(* IEC 61131-3 sources: JingjiangArm/moonboxpro_arm_8.4/Application/Application/任务列表/ExtTask/动作处理/动作处理 (part 2) *)

(* ---- KS_FB_GrpFetchIOCtrl.st ---- *)
(*@CES
Name=KS_FB_GrpFetchIOCtrl
Type=FunctionBlock
TypeGuid=6f9dac99-8de1-4efc-8465-68ac443b7d08
Guid=a7ec576d-c0a8-4898-9e79-82769fd09b46
HasDeclaration=True
HasImplementation=True
*)
{DECLARATION}
FUNCTION_BLOCK KS_FB_GrpFetchIOCtrl
VAR_INPUT
	i_xEn: BOOL;
	i_iGrpId: INT;
	i_pstStEvtReq: POINTER TO StEvtReq; (* 沿触发标志 *)
	i_pstStSysCfgStruct: POINTER TO StSysCfgStruct;
	i_pastStIOMap_Main_FE						: POINTER TO ARRAY [1..4] OF StIOMap_Main_FE;(*轴io数据区域|AB系*)
	i_pastStIOMap_Axis_FE					: POINTER TO ARRAY [1..MAX_UNIT_NUM] OF StIOMap_Axis_FE;(*轴io数据区域|`````````````````````````````````````````````*)
	i_pastStIOMap_Axis_Extra_FE				: POINTER TO ARRAY [1..MAX_UNIT_NUM] OF StIOMap_Axis_Extra_FE;
	i_pastStIOMap_UwRw_FE_Uw					: POINTER TO ARRAY [1..2] OF StIOMap_UwRw_FE;(*轴io数据区域|AB系*)
	i_pastStIOMap_UwRw_FE_Rw					: POINTER TO ARRAY [1..2] OF StIOMap_UwRw_FE;(*轴io数据区域|AB系*)

	i_iUMax: INT;(*最大色组*)
	i_dwEquipmentProf: DWORD;(*机型：bit20:双收双放bit21:A放B收*)
	i_xUseRealStationOnRingnet: BOOL;(*使用真实站点*)
	i_axLinkage: ARRAY [1..MAX_UNIT_NUM] OF BOOL;
	i_axThisUnitEna: ARRAY [1..MAX_UNIT_NUM] OF BOOL;
	i_axSwitchOn_CoatingPrn: ARRAY [1..MAX_UNIT_NUM] OF BOOL;

	i_xIsValid_If_I: BOOL;
	i_xIsValid_If_II: BOOL;
	i_xIsValid_Of_I: BOOL;
	i_xIsValid_Of_II: BOOL;
//	i_pstStRingInfVer1: POINTER TO StRingInfVer1; (* 所有站点列表 *)

	//2026.5.20.133000 by liu.yt 使用map生成的系统站信息列表@根据实际站生成
	//i_pstStStationInfo_KS: POINTER TO StStationInfo_KS;
	(*输出列表*)
	i_pstStSysStationInf	: POINTER TO StSysStationInf;
	i_pxInit_StationList	: POINTER TO BOOL;

END_VAR
VAR_OUTPUT
	o_xEn: BOOL;
	o_iErNo: INT;
	o_iGrpAxisNum_Pu: INT; (* 系的色组数量|色组按照从小到大排序了 *)
	o_iGrpAxisTotalNum: INT; (* 系的轴数量 *)
	o_aiGrpAxisList: ARRAY [1..MAX_UNIT_NUM] OF INT; (* 系的轴列表 *)
	o_iIOGrpIdx_Uw: INT; (* 放料id *)
	o_iIOGrpIdx_Rw: INT; (* 收料id *)
	o_iAxisId_If_IOMapUse: INT; (* 放牵轴id *)
	o_iAxisId_Of_IOMapUse: INT; (* 收牵轴id *)
	o_aiGrpServoAxisList_Uw: ARRAY [1..2] OF INT := [2(-1)]; (* 2021.5.7.150202/目前仅支持双工位/[1]放置A轴/[2]放置B轴/轴id(-1)表无效 *)
	o_aiGrpServoAxisList_Rw: ARRAY [1..2] OF INT := [2(-1)]; (* 2021.5.7.150202/目前仅支持双工位/[1]放置A轴/[2]放置B轴/轴id(-1)表无效 *)

	(*2022.5.25.103645 增加联动轴*)
	o_iGrpLinkageAxisNum_Pu: INT; (* 系的色组联动轴数量|色组按照从小到大排序了 *)
	o_aiGrpLinkageAxisList: ARRAY [1..MAX_UNIT_NUM] OF INT; (* 系的联动轴列表 *)
	(*2023.09.04.131040 增加了色序列表的输出*)
	o_iGrpArcAxisNum_Pu: INT; (* 系的色联动轴套色打开数量|色组按照从小到大排序了 *)
	o_aiGrpArcAxisList: ARRAY [1..MAX_UNIT_NUM] OF INT; (* 系的联动轴套色打开列表 *)
	o_aiGrpArcIdList: ARRAY [1..MAX_UNIT_NUM] OF INT; (* 系的联动轴套色Id列表@2024.02.22.083346 套色id有可能会手动修改 *)
	o_aiGrpFollowArcIdList: ARRAY [1..MAX_UNIT_NUM] OF INT; (* 系的联动轴套色跟踪色序Id列表@2024.02.22.083346 和套色个数同步更新*)

(*运动列表*)
	o_iAxisNum_Trap: INT;(*点位运动轴数量*)
	o_aiStationList_Trap: ARRAY [1..MAX_STATION_NUM] OF INT;(*点位运动轴列表*)
	o_iAxisNum_Gear: INT;(*电子齿轮运动轴数量*)
	o_aiStationList_Gear: ARRAY [1..MAX_STATION_NUM] OF INT;(*电子齿轮运动轴列表*)
	o_iAxisNum_GantrayTrap: INT;(*龙门点位运动组数量*)
	o_aiStationList_GantrayTrap: ARRAY [1..MAX_STATION_NUM] OF INT;(*龙门点位运动轴列表*)
	o_iAxisNum_Jog: INT;(*龙门点位运动组数量*)
	o_aiStationList_Jog: ARRAY [1..MAX_STATION_NUM] OF INT;(*龙门点位运动轴列表*)
	o_iAxisNum_All: INT;
	o_aiStationList_All: ARRAY [1..MAX_STATION_NUM] OF INT;
	o_aiIndexList_All_Trap: ARRAY [1..MAX_STATION_NUM] OF INT;(*点位运动轴列表*)
	o_aiIndexList_All_Gear: ARRAY [1..MAX_STATION_NUM] OF INT;(*电子齿轮运动轴列表*)
	o_aiIndexList_All_Gantray: ARRAY [1..MAX_STATION_NUM] OF INT;(*龙门点位运动轴列表*)
	o_aiIndexList_All_Jog: ARRAY [1..MAX_STATION_NUM] OF INT;(*龙门点位运动轴列表*)
	o_axFlag_SlaveUseCmm_Pro: ARRAY [1..MAX_UNIT_NUM] OF BOOL;(*色组使用PRO/月光宝盒*)
	//2026.04.10.145314
	o_dwAxisFlags_Estop:DWORD;(*系急停状态*)
END_VAR
VAR_IN_OUT
	io_abyColorIdCurrent: ARRAY [1..MAX_UNIT_NUM] OF BYTE;(*色组色序*)
	io_abyFollowColorId: ARRAY [1..MAX_UNIT_NUM] OF BYTE;
END_VAR
VAR
	iN: INT;
	iK: INT;
	iTmpAxisId: INT;
	afbR_TRIG_EvtReq: ARRAY [1..17] OF R_TRIG; (* 上升沿触发器 *)
	dwMaskMonitoring_Estop: DWORD; (* 急停标志位输出 *)
	dwMaskMonitoring_Stop: DWORD;
	dwMaskMonitoring_FastStop: DWORD;
	dwMaskMonitoring_Tension: DWORD;
	dwMaskMonitoring_ManuSpdUp: DWORD;
	dwMaskMonitoring_ManuSpdDn: DWORD;
	dwMaskMonitoring_Ink: DWORD;
	dwMaskMonitoring_Prestart: DWORD;
	dwMaskMonitoring_PressAll: DWORD;
	dwMaskMonitoring_UnpressAll: DWORD;
	dwMaskMonitoring_Print: DWORD;
	dwMaskMonitoring_AlarmBell: DWORD;
	dwMaskMonitoring_AllInchRun: DWORD;
	dwMaskMonitoring_AllExhBlower: DWORD;
	dwMaskMonitoring_AllCoolBlower: DWORD;
	dwMaskMonitoring_AllHotBlower: DWORD;
	dwMaskMonitoring_AllHeating: DWORD;
	xIsDualUwRw: BOOL := FALSE; (* 双收双放 *)
	xAsOneMachine: BOOL := FALSE; (* A放B收结构 *)
	iUnitId: INT;
	iGrpId: INT;
	iTypeId: INT;
	iAxisTypeId: INT;
	xInit_ColorId: BOOL;(*开机初始化一次色序ID*)
	byColorID: BYTE;
	pstStIOMap_AxisBasic: POINTER TO StIOMap_Axis_FE; (* 基础io *)
	pstStIOMap_AxisExtra: POINTER TO StIOMap_Axis_Extra_FE; (* 扩展io *)
	axArcEnSts_Bak:ARRAY [1..MAX_STATION_NUM] OF BOOL;
	abyArcId_Bak:ARRAY [1..MAX_STATION_NUM] OF BYTE;
	iUnitId_Rd: INT;
	iTypeId_Rd: INT;
	//iAxisId_Rd: INT;
	//iCoreId_Rd: INT;
	//iGroupId_Rd: INT;
	//iAdjAxisId_Rd: INT;

	//2026.5.20.133421 by liu.yt
	pstStationInf:POINTER TO StStationInf;//每个站的信息
END_VAR

{IMPLEMENTATION}
o_xEn:= i_xEn;
o_iErNo:= 0;

(* 返回值初始化 *)
o_iIOGrpIdx_Uw:= -1; (* 放料io系id初始化 *)
o_iIOGrpIdx_Rw:= -1; (* 收料io系id初始化 *)
o_iAxisId_If_IOMapUse:= -1; (* 放牵轴id初始化 *)
o_iAxisId_Of_IOMapUse:= -1; (* 收牵轴id初始化 *)
o_iGrpAxisNum_Pu:= 0; (* 输出色组数量初始化 *)
o_iGrpAxisTotalNum:= 0; (* 输出总轴数量初始化 *)
o_iGrpLinkageAxisNum_Pu:= 0; (* 输出联动色组数量初始化 *)
o_iGrpArcAxisNum_Pu:=0;
FOR iN:=1 TO MAX_UNIT_NUM BY 1 DO(* 轴列表初始化 *)
	o_aiGrpAxisList[iN]:= -1;
	o_aiGrpLinkageAxisList[iN]:= -1;
	o_aiGrpArcAxisList[iN]:=-1;
	o_aiGrpArcIdList[iN]:=-1;(*2024.02.22.083413*)
	o_aiGrpFollowArcIdList[iN]:=-1;
END_FOR
o_aiGrpServoAxisList_Uw[1]:= -1;
o_aiGrpServoAxisList_Uw[2]:= -1;

o_aiGrpServoAxisList_Rw[1]:= -1;
o_aiGrpServoAxisList_Rw[2]:= -1;

(* 2018.9.4.162654\增加的监控初始化 *)
dwMaskMonitoring_Estop:= 0;
dwMaskMonitoring_Stop:= 0;
dwMaskMonitoring_Tension:= 0;
dwMaskMonitoring_ManuSpdUp:= 0;
dwMaskMonitoring_ManuSpdDn:= 0;
dwMaskMonitoring_Ink:= 0;
dwMaskMonitoring_Prestart:= 0;
dwMaskMonitoring_PressAll:= 0;
dwMaskMonitoring_UnpressAll:= 0;
dwMaskMonitoring_Print:= 0;
dwMaskMonitoring_AlarmBell:= 0;
dwMaskMonitoring_AllInchRun:= 0;
dwMaskMonitoring_AllExhBlower:= 0;
dwMaskMonitoring_AllCoolBlower:= 0;
dwMaskMonitoring_AllHotBlower:= 0;
dwMaskMonitoring_AllHeating:= 0;

IF i_xEn THEN
	IF (i_iGrpId=1 OR i_iGrpId=2) AND
		i_pstStEvtReq<>0 AND
		i_pastStIOMap_Main_FE<>0 AND
		i_pastStIOMap_Axis_FE<>0 AND
		i_pastStIOMap_Axis_Extra_FE<>0 AND
		i_pastStIOMap_UwRw_FE_Uw<>0 AND
		i_pastStIOMap_UwRw_FE_Rw<>0 AND
		i_pxInit_StationList<>0 THEN
		KS_InitStEvtReq(i_pstStEvtReq); (* 初始化StEvtReq@2018.7.31.094400 *)
		xIsDualUwRw:= i_dwEquipmentProf.20;
		xAsOneMachine:= i_dwEquipmentProf.21;
		IF NOT(i_iUMax>=1 AND i_iUMax<=16) THEN
			o_iErNo:=-4;
			RETURN;
		END_IF
		IF xIsDualUwRw AND xAsOneMachine AND i_iGrpId<>1 THEN(* A放B收\操作了A系以外的系 *)
			o_iErNo:= -2;
			RETURN;
		ELSIF (NOT xIsDualUwRw) AND i_iGrpId<>1 THEN(* 对于标准机型操作了A系以外的系 *)
			o_iErNo:= -3;
			RETURN;
		ELSE(* 其余正常情况 *)
			(* 生成当前系数的色组轴号列表|
			/*目前1个系内的放牵和收牵只认为各有1个,所以读取轴类型是牵引的会覆盖前面的取值 *)
			IF i_xUseRealStationOnRingnet THEN
// 				FOR iN:=1 TO i_pstStStationInfo_KS^.iStationNum BY 1 DO
// 					KS_GetAxisIdForMotByStation_V2(
// 						i_iStationId:= i_pstStStationInfo_KS^.aiStationId_List[iN],
// 						i_piAxisId:= ADR(iAxisId_Rd),
// 						i_piTypeId:= ADR(iTypeId_Rd),
// 						i_piUnitId:= ADR(iUnitId_Rd),
// 						i_piCoreId:= ADR(iCoreId_Rd),
// 						i_piGroupId:= ADR(iGroupId_Rd),
// 						i_piAdjAxisId:= ADR(iAdjAxisId_Rd),
// 						i_pstStSysStationInf:= ADR(g_stStSysStationInf));
// 					IF iUnitId_Rd>=1 AND iUnitId<=MAX_UNIT_NUM THEN
// 						iGrpId:= KS_GetGrpIdByAxisId(iUnitId,ADR(g_stStSysParam),ADR(iAxisTypeId));
// 						//2026.5.12.112929就用版辊驱动器数量输出轴列表吧
// 						IF iGrpId= i_iGrpId THEN
// 							IF iTypeId_Rd=TYPE_UNIT_PRN THEN
// 								o_iGrpAxisNum_Pu:= o_iGrpAxisNum_Pu+1;
// 								o_aiGrpAxisList[o_iGrpAxisNum_Pu]:= iUnitId_Rd;
// 							END_IF
// 						END_IF
// 					END_IF
// 				END_FOR
				//2026.5.20.133216 by liu.yt 重新生成列表@根据实际站
				FOR iN:=1 TO BYTE_TO_INT(i_pstStSysStationInf^.byStationNum) BY 1 DO
					pstStationInf:=ADR(i_pstStSysStationInf^.astStationInf[iN]);

					KS_GetAxisIdForMotByStation_V2(
						i_iStationId:= pstStationInf^.iStationId,
						i_piAxisId:= 0,
						i_piTypeId:= ADR(iTypeId_Rd),
						i_piUnitId:= ADR(iUnitId_Rd),
						i_piCoreId:= 0,
						i_piGroupId:= 0,
						i_piAdjAxisId:= 0,
						i_pstStSysStationInf:= i_pstStSysStationInf);
					IF iUnitId_Rd>=1 AND iUnitId_Rd<=MAX_UNIT_NUM THEN//色组id合法@1个色组可能会存在多个不同功能站号返回。我们只检查色组轴
						iGrpId:= KS_GetGrpIdByAxisId(iUnitId_Rd,ADR(g_stStSysParam),ADR(iAxisTypeId));
						//2026.5.12.112929就用版辊驱动器数量输出轴列表吧
						IF iGrpId= i_iGrpId THEN
							IF iTypeId_Rd=TYPE_UNIT_CTL THEN
								o_iGrpAxisNum_Pu:= o_iGrpAxisNum_Pu+1;
								o_aiGrpAxisList[o_iGrpAxisNum_Pu]:= iUnitId_Rd;
							END_IF
						END_IF
					END_IF
				END_FOR
			ELSE
				(* 2020.9.11.134731
				** 按照系统配置的色组填充列表|
				** *)
				FOR iUnitId:=1 TO i_iUMax BY 1 DO
					o_iGrpAxisNum_Pu:= o_iGrpAxisNum_Pu+1;
					o_aiGrpAxisList[o_iGrpAxisNum_Pu]:= iUnitId;
				END_FOR
			END_IF

			(* **
			** 将牵引轴使能出来@2019.4.26.171841
			** 针对给了使能|但没有给牵引指定一个有效的轴id
			** *)
			IF NOT xIsDualUwRw THEN(* 非双收双放 *)
				(* 放牵轴id *)
				IF i_xIsValid_If_I THEN
					o_iAxisId_If_IOMapUse:= 1;
				END_IF

				(* 收牵轴id *)
				IF i_xIsValid_Of_I THEN
					o_iAxisId_Of_IOMapUse:= 2;
				END_IF
			ELSE(* 双收双放 *)
				IF xAsOneMachine THEN(* A放B收 *)
					IF i_iGrpId=1 THEN
						(* 放牵轴id *)
						IF i_xIsValid_If_I THEN
							o_iAxisId_If_IOMapUse:= 1;
						END_IF

						(* 收牵轴id *)
						IF i_xIsValid_Of_II THEN
							o_iAxisId_Of_IOMapUse:= 4;
						END_IF
					END_IF
				ELSE(* A放A收|B放B收 *)
					IF i_iGrpId=1 THEN
						(* 放牵轴id *)
						IF i_xIsValid_If_I THEN
							o_iAxisId_If_IOMapUse:= 1;
						END_IF

						(* 收牵轴id *)
						IF i_xIsValid_Of_I THEN
							o_iAxisId_Of_IOMapUse:= 2;
						END_IF
					ELSE(* B系 *)
						(* 放牵轴id *)
						IF i_xIsValid_If_II THEN
							o_iAxisId_If_IOMapUse:= 3;
						END_IF

						(* 收牵轴id *)
						IF i_xIsValid_Of_II THEN
							o_iAxisId_Of_IOMapUse:= 4;
						END_IF
					END_IF
				END_IF
			END_IF
			(* 色组按从小到大的编号排列 *)
			FOR iN:=o_iGrpAxisNum_Pu TO 2 BY -1 DO
				FOR iK:=1 TO iN BY 1 DO
					IF o_aiGrpAxisList[iN]<o_aiGrpAxisList[iK] THEN
						iTmpAxisId:= o_aiGrpAxisList[iN];
						o_aiGrpAxisList[iN]:= o_aiGrpAxisList[iK];
						o_aiGrpAxisList[iK]:= iTmpAxisId;
					END_IF
				END_FOR
			END_FOR

			(* 在色组轴号之后追加牵引轴编号 *)
			o_iGrpAxisTotalNum:= o_iGrpAxisNum_Pu;
(*2026.5.12.132915这个列表只放色组相关的
			(* 放牵 *)
			IF o_iAxisId_If_IOMapUse>=1 AND o_iAxisId_If_IOMapUse<=MAX_STATION_NUM THEN
				o_iGrpAxisTotalNum:= o_iGrpAxisTotalNum+1;
				o_aiGrpAxisList[o_iGrpAxisTotalNum]:= o_iAxisId_If_IOMapUse;
			END_IF

			(* 收牵 *)
			IF o_iAxisId_Of_IOMapUse>=1 AND o_iAxisId_Of_IOMapUse<=MAX_STATION_NUM THEN
				o_iGrpAxisTotalNum:= o_iGrpAxisTotalNum+1;
				o_aiGrpAxisList[o_iGrpAxisTotalNum]:= o_iAxisId_Of_IOMapUse;
			END_IF
*)
			(*2022.5.25.104049 增加联动轴的列表输出*)
			FOR iN:=1 TO o_iGrpAxisNum_Pu BY 1 DO
				iTmpAxisId:= o_aiGrpAxisList[iN];
				IF iTmpAxisId>0 THEN
					IF i_axLinkage[iTmpAxisId] THEN(*联动*)
						o_iGrpLinkageAxisNum_Pu:=o_iGrpLinkageAxisNum_Pu+1;
						o_aiGrpLinkageAxisList[o_iGrpLinkageAxisNum_Pu]:=iTmpAxisId;
					END_IF
				END_IF
			END_FOR

			(*2023.09.04.131214 增加联动轴套色打开的列表输出*)
			IF xInit_ColorId THEN
				FOR iN:=1 TO o_iGrpLinkageAxisNum_Pu BY 1 DO
					iTmpAxisId:= o_aiGrpLinkageAxisList[iN];
					IF iTmpAxisId>0 THEN
						IF io_abyColorIdCurrent[iTmpAxisId]>0 AND io_abyColorIdCurrent[iTmpAxisId]<=MAX_UNIT_NUM THEN(*色序合法*)
							o_iGrpArcAxisNum_Pu:=o_iGrpArcAxisNum_Pu+1;
							o_aiGrpArcAxisList[o_iGrpArcAxisNum_Pu]:=iTmpAxisId;
							o_aiGrpArcIdList[o_iGrpArcAxisNum_Pu]:=io_abyColorIdCurrent[iTmpAxisId];(*2024.02.22.083448 套色id也统计出来*)
							o_aiGrpFollowArcIdList[o_iGrpArcAxisNum_Pu]:=io_abyFollowColorId[iTmpAxisId];(*2024.02.22.112812 界面修改或者一些开关控制*)
						END_IF
					END_IF
				END_FOR
			END_IF

			IF xIsDualUwRw THEN
				(* 双收双放 *)

				IF xAsOneMachine THEN
					(* A放B收 *)
					o_iIOGrpIdx_Uw:= 1;
					o_iIOGrpIdx_Rw:= 2;
				ELSE
					(* A/B系各自用各自的 *)
					IF i_iGrpId=1 THEN
						o_iIOGrpIdx_Uw:= 1;
						o_iIOGrpIdx_Rw:= 1;
					ELSE
						o_iIOGrpIdx_Uw:= 2;
						o_iIOGrpIdx_Rw:= 2;
					END_IF
				END_IF
			ELSE(* 普通机型\只看A系 *)
				o_iIOGrpIdx_Uw:= 1;
				o_iIOGrpIdx_Rw:= 1;
			END_IF

			(* 放料和收料的急停按钮 *)
			IF i_pastStIOMap_UwRw_FE_Uw^[o_iIOGrpIdx_Uw].i_xEstop THEN(* 放料急停 *)
				dwMaskMonitoring_Estop:= dwMaskMonitoring_Estop OR SHL(DWORD#1,20);
				i_pstStEvtReq^.xEvt_Estop:= TRUE;
			END_IF
			IF i_pastStIOMap_UwRw_FE_Rw^[o_iIOGrpIdx_Rw].i_xEstop THEN(* 收料急停 *)
				dwMaskMonitoring_Estop:= dwMaskMonitoring_Estop OR SHL(DWORD#1,21);
				i_pstStEvtReq^.xEvt_Estop:= TRUE;
			END_IF

			(*放牵收牵的按钮处理*)
			IF i_pastStIOMap_Main_FE^[o_iAxisId_If_IOMapUse].i_xEstop OR
				i_pastStIOMap_Main_FE^[o_iAxisId_Of_IOMapUse].i_xEstop THEN
				i_pstStEvtReq^.xEvt_Estop:= TRUE;
			END_IF
			IF i_pastStIOMap_Main_FE^[o_iAxisId_If_IOMapUse].i_xStop OR
				i_pastStIOMap_Main_FE^[o_iAxisId_Of_IOMapUse].i_xStop THEN
				i_pstStEvtReq^.xEvt_Stop:= TRUE;
			END_IF
			IF i_pastStIOMap_Main_FE^[o_iAxisId_If_IOMapUse].i_xFastStop OR
				i_pastStIOMap_Main_FE^[o_iAxisId_Of_IOMapUse].i_xFastStop THEN
				//2026.06.04.145510 变量写错了 by liu.yt
				//i_pstStEvtReq^.xEvt_Stop:= TRUE;
				i_pstStEvtReq^.xEvt_FastStop:= TRUE;
			END_IF
			IF i_pastStIOMap_Main_FE^[o_iAxisId_If_IOMapUse].i_xTension OR
				i_pastStIOMap_Main_FE^[o_iAxisId_Of_IOMapUse].i_xTension THEN
				i_pstStEvtReq^.xEvt_Tension:= TRUE;
			END_IF
			IF i_pastStIOMap_Main_FE^[o_iAxisId_If_IOMapUse].i_xAcc OR
				i_pastStIOMap_Main_FE^[o_iAxisId_Of_IOMapUse].i_xAcc THEN
				i_pstStEvtReq^.xEvt_ManuSpdUp:= TRUE;
			END_IF
			IF i_pastStIOMap_Main_FE^[o_iAxisId_If_IOMapUse].i_xDec OR
				i_pastStIOMap_Main_FE^[o_iAxisId_Of_IOMapUse].i_xDec THEN
				i_pstStEvtReq^.xEvt_ManuSpdDn:= TRUE;
			END_IF
			IF i_pastStIOMap_Main_FE^[o_iAxisId_If_IOMapUse].i_xInk OR
				i_pastStIOMap_Main_FE^[o_iAxisId_Of_IOMapUse].i_xInk THEN
				i_pstStEvtReq^.xEvt_Ink:= TRUE;
			END_IF
			IF i_pastStIOMap_Main_FE^[o_iAxisId_If_IOMapUse].i_xPrestart OR
				i_pastStIOMap_Main_FE^[o_iAxisId_Of_IOMapUse].i_xPrestart THEN
				i_pstStEvtReq^.xEvt_Prestart:= TRUE;
			END_IF
			IF i_pastStIOMap_Main_FE^[o_iAxisId_If_IOMapUse].i_xPrint OR
				i_pastStIOMap_Main_FE^[o_iAxisId_Of_IOMapUse].i_xPrint THEN
				i_pstStEvtReq^.xEvt_Print:= TRUE;
			END_IF
			IF i_pastStIOMap_Main_FE^[o_iAxisId_If_IOMapUse].i_xPressAll OR
				i_pastStIOMap_Main_FE^[o_iAxisId_Of_IOMapUse].i_xPressAll THEN
				i_pstStEvtReq^.xEvt_PressAll:= TRUE;
			END_IF
			IF i_pastStIOMap_Main_FE^[o_iAxisId_If_IOMapUse].i_xUnPressAll OR
				i_pastStIOMap_Main_FE^[o_iAxisId_Of_IOMapUse].i_xUnPressAll THEN
				i_pstStEvtReq^.xEvt_UnPressAll:= TRUE;
			END_IF
			IF i_pastStIOMap_Main_FE^[o_iAxisId_If_IOMapUse].i_xAlarmBell OR
				i_pastStIOMap_Main_FE^[o_iAxisId_Of_IOMapUse].i_xAlarmBell THEN
				i_pstStEvtReq^.xEvt_AlarmBell:= TRUE;
			END_IF

			IF i_pastStIOMap_Main_FE^[o_iAxisId_If_IOMapUse].i_xAllExhBlower_Up OR
				i_pastStIOMap_Main_FE^[o_iAxisId_Of_IOMapUse].i_xAllExhBlower_Up OR
				i_pastStIOMap_Main_FE^[o_iAxisId_If_IOMapUse].i_xAllExhBlower_Dn OR
				i_pastStIOMap_Main_FE^[o_iAxisId_Of_IOMapUse].i_xAllExhBlower_Dn THEN
				(* 整机排风 *)
				i_pstStEvtReq^.xEvt_AllExhBlower:= TRUE;
			END_IF

			IF i_pastStIOMap_Main_FE^[o_iAxisId_If_IOMapUse].i_xAllCoolBlower OR
				i_pastStIOMap_Main_FE^[o_iAxisId_Of_IOMapUse].i_xAllCoolBlower THEN
				(* 整机冷风 *)
				i_pstStEvtReq^.xEvt_AllCoolBlower:= TRUE;
			END_IF
			IF i_pastStIOMap_Main_FE^[o_iAxisId_If_IOMapUse].i_xAllHotBlower OR
				i_pastStIOMap_Main_FE^[o_iAxisId_Of_IOMapUse].i_xAllHotBlower THEN
				(* 整机热风 *)
				i_pstStEvtReq^.xEvt_AllHotBlower:= TRUE;
			END_IF
			IF i_pastStIOMap_Main_FE^[o_iAxisId_If_IOMapUse].i_xAllHeating OR
				i_pastStIOMap_Main_FE^[o_iAxisId_Of_IOMapUse].i_xAllHeating THEN
				(* 整机加热 *)
				i_pstStEvtReq^.xEvt_AllHeating:= TRUE;
			END_IF

			(* 默认3档开关 作互斥 *)
			IF i_pastStIOMap_Main_FE^[o_iAxisId_Of_IOMapUse].i_xTapPosition_Breaking THEN(* 2018.7.16.151749\断料档位 *)
				i_pstStEvtReq^.xEvt_TapPosition_Breaking:= TRUE;
				i_pstStEvtReq^.xEvt_TapPosition_UniformInk:= FALSE;
				i_pstStEvtReq^.xEvt_TapPosition_Printing:= FALSE;
			ELSIF i_pastStIOMap_Main_FE^[o_iAxisId_Of_IOMapUse].i_xTapPosition_UniformInk THEN(* 2018.7.16.152023\匀墨档位 *)
				i_pstStEvtReq^.xEvt_TapPosition_UniformInk:= TRUE;
				i_pstStEvtReq^.xEvt_TapPosition_Breaking:= FALSE;
				i_pstStEvtReq^.xEvt_TapPosition_Printing:= FALSE;
			ELSE(* 2018.7.16.152128\印刷档位 *)
				i_pstStEvtReq^.xEvt_TapPosition_Printing:= TRUE;
				i_pstStEvtReq^.xEvt_TapPosition_Breaking:= FALSE;
				i_pstStEvtReq^.xEvt_TapPosition_UniformInk:= FALSE;
			END_IF

			(* 影响整机的逻辑按钮\所有轴上可能都有\就在FOR循环里面检查(当然要包含牵引) *)
			byColorID:=0;(*2022.6.8.101746*)
			FOR iN:=1 TO o_iGrpAxisNum_Pu BY 1 DO
				iUnitId:= o_aiGrpAxisList[iN]; (* 列表由于本地生成\所以iAxisId可以不检查 *)
				pstStIOMap_AxisBasic:= ADR(i_pastStIOMap_Axis_FE^[iUnitId]); (* 基础io表 *)
				pstStIOMap_AxisExtra:= ADR(i_pastStIOMap_Axis_Extra_FE^[iUnitId]); (* 扩展io表 *)

				IF pstStIOMap_AxisBasic^.i_xEstop THEN
					(* 急停 *)
					i_pstStEvtReq^.xEvt_Estop:= TRUE;
					dwMaskMonitoring_Estop:= dwMaskMonitoring_Estop OR SHL(DWORD#1,iUnitId-1);
				END_IF
				IF pstStIOMap_AxisBasic^.i_xStop THEN
					(* 停机 *)
					i_pstStEvtReq^.xEvt_Stop:= TRUE;
					dwMaskMonitoring_Stop:= dwMaskMonitoring_Stop OR SHL(DWORD#1,iUnitId-1);
				END_IF

				IF pstStIOMap_AxisBasic^.i_xAcc THEN
					(* 手动加速 *)
					i_pstStEvtReq^.xEvt_ManuSpdUp:= TRUE;
					dwMaskMonitoring_ManuSpdUp:= dwMaskMonitoring_ManuSpdUp OR SHL(DWORD#1,iUnitId-1);
				END_IF
				IF pstStIOMap_AxisBasic^.i_xDec THEN
					(* 手动减速 *)
					i_pstStEvtReq^.xEvt_ManuSpdDn:= TRUE;
					dwMaskMonitoring_ManuSpdDn:= dwMaskMonitoring_ManuSpdDn OR SHL(DWORD#1,iUnitId-1);
				END_IF

				IF pstStIOMap_AxisBasic^.i_xAlarmBell THEN
					(* 警铃 *)
					i_pstStEvtReq^.xEvt_AlarmBell:= TRUE;
					dwMaskMonitoring_AlarmBell:= dwMaskMonitoring_AlarmBell OR SHL(DWORD#1,iUnitId-1);
				END_IF
				IF pstStIOMap_AxisBasic^.i_xInch AND
					i_axLinkage[iUnitId] THEN
					(* 整机单运行 *)
					i_pstStEvtReq^.xEvt_AllInchRun:= TRUE;
					dwMaskMonitoring_AllInchRun:= dwMaskMonitoring_AllInchRun OR SHL(DWORD#1,iUnitId-1);
				END_IF
			END_FOR

			//2026.5.9.172930
			//2026.04.10.145142 + 系急停变量赋值
			o_dwAxisFlags_Estop:=dwMaskMonitoring_Estop;

			(*2024.02.21.084550 优化套色id逻辑*)
			KS_GetArcIdList(
				TRUE(*i_xEn*),
				o_iGrpAxisNum_Pu(*i_iGrpAxisNum_Pu*),
				o_aiGrpAxisList(*i_aiGrpAxisList*),
				ADR(axArcEnSts_Bak)(*i_paxArcEnSts_Bak*),
				ADR(abyArcId_Bak)(*i_pabyArcId_Bak*),
				0(*i_piGrpArcAxisNum_Pu*),
				i_axLinkage,
				i_axThisUnitEna,
				i_axSwitchOn_CoatingPrn,
				ADR(io_abyColorIdCurrent));
			xInit_ColorId:=TRUE;

		END_IF

		(*2025.6.16.165421运动所有的轴列表处理一下*)
		IF NOT i_pxInit_StationList^ THEN
			i_pxInit_StationList^:= TRUE;
			o_iAxisNum_Trap:= 0;
			o_iAxisNum_Gear:= 0;
			o_iAxisNum_GantrayTrap:= 0;
			o_iAxisNum_Jog:= 0;
			o_iAxisNum_All:= 0;
			FOR iN:=1 TO MAX_STATION_NUM BY 1 DO
				o_aiStationList_Trap[iN]:= 0;
				o_aiStationList_Gear[iN]:= 0;
				o_aiStationList_GantrayTrap[iN]:= 0;
				o_aiStationList_All[iN]:= 0;
				o_aiIndexList_All_Trap[iN]:= 0;
				o_aiIndexList_All_Gear[iN]:= 0;
				o_aiIndexList_All_Gantray[iN]:= 0;
			END_FOR

			FOR iN:=1 TO i_pstStSysStationInf^.byStationNum BY 1 DO
				pstStationInf:=ADR(i_pstStSysStationInf^.astStationInf[iN]);
				KS_GetUnitIdAndTypeByStationId(
					pstStationInf^.iStationId ,//i_pstStRingInfVer1^.m_station_id_list[iN],//i_pstStStationInfo_KS^.aiStationId_List[iN], //,
					ADR(iUnitId),
					ADR(iTypeId),
					i_pstStSysCfgStruct);
				IF iTypeId= OBJ_IS_HORIZ_MOTION OR
					 iTypeId=OBJ_IS_PHOTOCELL THEN(*光电眼行走机构 | 2024.04.01.092649*)
					o_iAxisNum_Trap:= o_iAxisNum_Trap+1;
					IF o_iAxisNum_Trap<>0 THEN
						o_aiStationList_Trap[o_iAxisNum_Trap]:= pstStationInf^.iStationId;//i_pstStRingInfVer1^.m_station_id_list[iN];//
						o_aiIndexList_All_Trap[o_iAxisNum_Trap]:= iN;
					END_IF
				ELSIF iTypeId= OBJ_IS_PRN_ROLLER_PRESSURE_M OR
					iTypeId= OBJ_IS_PRN_ROLLER_PRESSURE_G OR
					iTypeId= OBJ_IS_NET_ROLLER_PRESSURE_M OR
					iTypeId= OBJ_IS_NET_ROLLER_PRESSURE_G OR
					iTypeId= OBJ_IS_STR_ROLLER_PRESSURE_M OR
					iTypeId= OBJ_IS_STR_ROLLER_PRESSURE_G THEN
					o_iAxisNum_GantrayTrap:= o_iAxisNum_GantrayTrap+1;
					IF o_iAxisNum_GantrayTrap<>0 THEN
						o_aiStationList_GantrayTrap[o_iAxisNum_GantrayTrap]:= pstStationInf^.iStationId;//i_pstStRingInfVer1^.m_station_id_list[iN];//;
						o_aiIndexList_All_Gantray[o_iAxisNum_GantrayTrap]:= iN;

					END_IF
				ELSIF iTypeId= OBJ_IS_UNWIND_A OR
					iTypeId= OBJ_IS_UNWIND_B OR
					iTypeId= OBJ_IS_REWIND_A OR
					iTypeId= OBJ_IS_REWIND_B OR
					iTypeId= OBJ_IS_INFEED OR
					iTypeId= OBJ_IS_OUTFEED OR
					iTypeId= OBJ_IS_BOTTOM_ROLLER OR
					iTypeId= OBJ_IS_PRN_ROLLER OR
					iTypeId= OBJ_IS_NET_ROLLER OR
					iTypeId= OBJ_IS_CENTRAL_DRUM THEN
					o_iAxisNum_Gear:= o_iAxisNum_Gear+1;
					IF o_iAxisNum_Gear<>0 THEN
						o_aiStationList_Gear[o_iAxisNum_Gear]:= pstStationInf^.iStationId;//i_pstStRingInfVer1^.m_station_id_list[iN];//;
						o_aiIndexList_All_Gear[o_iAxisNum_Gear]:= iN;

					END_IF

					//2026.05.08.141028 | + | 增加收放料伺服的标志
					IF iTypeId= OBJ_IS_UNWIND_A OR
						iTypeId= OBJ_IS_UNWIND_B OR
						iTypeId= OBJ_IS_REWIND_A OR
						iTypeId= OBJ_IS_REWIND_B THEN
						g_xUwRwIsServo := TRUE;
					END_IF
				//这部分的代码处理会有问题@2026.5.20.140553 by liu.yt
				ELSIF pstStationInf^.iStationId>=1
					AND pstStationInf^.iStationId<16
					AND (pstStationInf^.udiStationType=HY_YTPE_CMM_CR_PRO
					OR	pstStationInf^.udiStationType=HY_YTPE_CMM_CR) THEN//色组使用月光宝盒/PRO通讯
					IF pstStationInf^.udiStationType=HY_YTPE_CMM_CR_PRO THEN
						o_axFlag_SlaveUseCmm_Pro[pstStationInf^.iStationId]:= TRUE;
					ELSE
						o_axFlag_SlaveUseCmm_Pro[pstStationInf^.iStationId]:= FALSE;
					END_IF
				END_IF
				IF iTypeId= OBJ_IS_HORIZ_MOTION OR
					iTypeId= OBJ_IS_PRN_ROLLER_PRESSURE_M OR
					iTypeId= OBJ_IS_PRN_ROLLER_PRESSURE_G OR
					iTypeId= OBJ_IS_NET_ROLLER_PRESSURE_M OR
					iTypeId= OBJ_IS_NET_ROLLER_PRESSURE_G OR
					iTypeId= OBJ_IS_UNWIND_A OR
					iTypeId= OBJ_IS_UNWIND_B OR
					iTypeId= OBJ_IS_REWIND_A OR
					iTypeId= OBJ_IS_REWIND_B OR
					iTypeId= OBJ_IS_INFEED OR
					iTypeId= OBJ_IS_OUTFEED OR
					iTypeId= OBJ_IS_BOTTOM_ROLLER OR
					iTypeId= OBJ_IS_PRN_ROLLER OR
					iTypeId= OBJ_IS_NET_ROLLER OR
					iTypeId= OBJ_IS_CENTRAL_DRUM OR//所有参与运动的轴个数
					iTypeId= OBJ_IS_PHOTOCELL OR
					iTypeId= OBJ_IS_STR_ROLLER_PRESSURE_M OR
					iTypeId= OBJ_IS_STR_ROLLER_PRESSURE_G THEN//所有参与运动的轴个数
					o_iAxisNum_All:= o_iAxisNum_All+1;
					IF o_iAxisNum_All<>0 THEN
						o_aiStationList_All[o_iAxisNum_All]:= pstStationInf^.iStationId;//i_pstStRingInfVer1^.m_station_id_list[iN];//;
					END_IF
				END_IF
			END_FOR
		END_IF

		(*-----------end--------------------------*)

		(* 上升沿检测 *)
		afbR_TRIG_EvtReq[1](CLK:= i_pstStEvtReq^.xEvt_Estop, Q=> i_pstStEvtReq^.xReqEstop); (* 急停 *)
		afbR_TRIG_EvtReq[2](CLK:= i_pstStEvtReq^.xEvt_Stop, Q=> i_pstStEvtReq^.xReqStop); (* 停机 *)
		afbR_TRIG_EvtReq[3](CLK:= i_pstStEvtReq^.xEvt_Tension, Q=> i_pstStEvtReq^.xReqTension); (* 张力投入 *)
		afbR_TRIG_EvtReq[4](CLK:= i_pstStEvtReq^.xEvt_ManuSpdUp, Q=> i_pstStEvtReq^.xReqManuSpdUp); (* 手动加速|按着才加速 *)
		afbR_TRIG_EvtReq[5](CLK:= i_pstStEvtReq^.xEvt_ManuSpdDn, Q=> i_pstStEvtReq^.xReqManuSpdDn); (* 手动减速|按着才减速 *)
		afbR_TRIG_EvtReq[6](CLK:= i_pstStEvtReq^.xEvt_Ink, Q=> i_pstStEvtReq^.xReqInk); (* 空转 *)
		afbR_TRIG_EvtReq[7](CLK:= i_pstStEvtReq^.xEvt_Prestart, Q=> i_pstStEvtReq^.xReqPrestart); (* 启动|预备 *)
		afbR_TRIG_EvtReq[8](CLK:= i_pstStEvtReq^.xEvt_PressAll, Q=> i_pstStEvtReq^.xReqPressAll); (* 全体合压 *)
		afbR_TRIG_EvtReq[9](CLK:= i_pstStEvtReq^.xEvt_UnpressAll, Q=> i_pstStEvtReq^.xReqUnpressAll); (* 全体离压 *)
		afbR_TRIG_EvtReq[10](CLK:= i_pstStEvtReq^.xEvt_Print, Q=> i_pstStEvtReq^.xReqPrint); (* 印刷|联动 *)
		afbR_TRIG_EvtReq[11](CLK:= i_pstStEvtReq^.xEvt_AlarmBell, Q=> i_pstStEvtReq^.xReqAlarmBell); (* 警铃|按着才响 *)
		afbR_TRIG_EvtReq[12](CLK:= i_pstStEvtReq^.xEvt_AllInchRun, Q=> i_pstStEvtReq^.xReqAllInchRun); (* 整机单运行 *)
		afbR_TRIG_EvtReq[13](CLK:= i_pstStEvtReq^.xEvt_AllExhBlower, Q=> i_pstStEvtReq^.xReqAllExhBlower); (* 排风启动 *)
		afbR_TRIG_EvtReq[14](CLK:= i_pstStEvtReq^.xEvt_AllCoolBlower, Q=> i_pstStEvtReq^.xReqAllCoolBlower); (* 冷风启动 *)
		afbR_TRIG_EvtReq[15](CLK:= i_pstStEvtReq^.xEvt_AllHotBlower, Q=> i_pstStEvtReq^.xReqAllHotBlower); (* 热风启动 *)
		afbR_TRIG_EvtReq[16](CLK:= i_pstStEvtReq^.xEvt_AllHeating, Q=> i_pstStEvtReq^.xReqAllHeating); (* 加热启动 *)
		afbR_TRIG_EvtReq[17](CLK:= i_pstStEvtReq^.xEvt_FastStop, Q=> i_pstStEvtReq^.xReqFastStop); (* 快停按钮 *)
		(*记录日志和变频报警处理稍后*)
	END_IF
END_IF

(* ---- KS_FB_GrpIndicatorLampCtrl.st ---- *)
(*@CES
Name=KS_FB_GrpIndicatorLampCtrl
Type=FunctionBlock
TypeGuid=6f9dac99-8de1-4efc-8465-68ac443b7d08
Guid=046cf0cb-05a3-4565-9599-869039b6c2cc
HasDeclaration=True
HasImplementation=True
*)
{DECLARATION}
FUNCTION_BLOCK KS_FB_GrpIndicatorLampCtrl
VAR_INPUT
	i_xEn: BOOL;
	i_iGrpId:INT;
	i_iCustomerNameId:INT;
	i_iGrpAxisNum_PU: INT;
	i_aiGrpAxisList: ARRAY [1..MAX_UNIT_NUM] OF INT;
	i_pstStSysParam: POINTER TO StSysParam;
	i_pastStIOMap_AxisBasic: POINTER TO ARRAY [1..MAX_UNIT_NUM] OF StIOMap_Axis_FE;
	i_pastStIOMap_Main: POINTER TO ARRAY [1..4] OF StIOMap_Main_FE;(*基础io|*)
	i_iAxisId_If: INT;
	i_iAxisId_Of: INT;
END_VAR
VAR_OUTPUT
	o_xEno: BOOL;
	o_iErNo: INT;
END_VAR
VAR
	iN: INT;
	iAxisId: INT;
	pstStIOMap_AxisBasic: POINTER TO StIOMap_Axis_FE;
	pstStIOMap_Main: POINTER TO StIOMap_Main_FE;
	pstStIOMap_Main_If: POINTER TO StIOMap_Main_FE;
	pstStIOMap_Main_Of: POINTER TO StIOMap_Main_FE;
	tmNow: TIME;
	tmLastStateChanged_print: TIME;
	tmLastStateChanged_prestart: TIME; (* 2021.3.3.113856/上次状态改变的时间 *)
	tmLastStateChanged_Stop: TIME; (* 2022.4.10.001512/上次状态改变的时间 *)
	xLamp_Stop: BOOL;(*停止灯指示*)
END_VAR

{IMPLEMENTATION}
o_xEno:= i_xEn;
o_iErNo:= 0;
IF i_xEn THEN
	IF (i_iGrpAxisNum_PU>=0 AND i_iGrpAxisNum_PU<=MAX_UNIT_NUM) AND(*色组有效|*)
		i_pastStIOMap_AxisBasic<>0 THEN(*轴IO有效|*)

		tmNow:= TIME(); (* 2021.3.3.114019/ *)

		(*2022.4.9.225300 增加了停止时候停止指示灯的闪烁指示*)
		IF i_pstStSysParam^.astStGrpParam_UnSave[i_iGrpId].xFlag_Stoping  (*OR (*停止中|*)
			 i_pstStGrpParam^.xFlag_FastStoping*) THEN(*快速停止中*)
			IF tmNow-tmLastStateChanged_Stop>=T#200MS THEN
				xLamp_Stop:=NOT xLamp_Stop;(**)
				tmLastStateChanged_Stop:= tmNow; (* 2021.3.3.114723/ *)
			END_IF
		ELSE
			xLamp_Stop:=i_pstStSysParam^.astStGrpParam_UnSave[i_iGrpId].xFlag_Stop;
			tmLastStateChanged_Stop:= tmNow; (* 2021.3.3.114723/ *)
		END_IF

		FOR iN:=1 TO i_iGrpAxisNum_PU BY 1 DO
			iAxisId:= i_aiGrpAxisList[iN];
			IF iAxisId>=1 AND iAxisId<=MAX_UNIT_NUM THEN
				pstStIOMap_AxisBasic:=ADR(i_pastStIOMap_AxisBasic^[iAxisId]);(*读取轴IO|*)
				//pstStIOMap_Main_If:=ADR(i_pastStIOMap_Main^[i_iAxisId_If]);(*读取牵引轴IO|*)
				//pstStIOMap_Main_Of:=ADR(i_pastStIOMap_Main^[i_iAxisId_Of]);(*读取牵引轴IO|*)
				pstStIOMap_AxisBasic^.o_xLamp_Estop:= i_pstStSysParam^.astStGrpParam_UnSave[i_iGrpId].xFlag_Estop AND pstStIOMap_AxisBasic^.i_xEstop;(*急停灯输出|*)
				pstStIOMap_AxisBasic^.o_xLamp_Stop:= xLamp_Stop OR
												(NOT i_pstStSysParam^.astStUnitParam_Save[iAxisId].xLinkage AND NOT i_pstStSysParam^.astStGrpParam_UnSave[i_iGrpId].xFlag_Estop);(*停止灯输出|*)
				pstStIOMap_AxisBasic^.o_xLamp_Inch:= (i_pstStSysParam^.astStGrpParam_UnSave[i_iGrpId].xFlag_Ink OR i_pstStSysParam^.astStGrpParam_UnSave[i_iGrpId].xFlag_Print) AND (i_pstStSysParam^.astStUnitParam_Save[iAxisId].xLinkage);(*联动状态下空转或印刷|*)
				pstStIOMap_AxisBasic^.o_xLamp_AxisError:= (i_pstStSysParam^.astStUnitParam_UnSave[iAxisId].xNetOffline_PrnRoller OR i_pstStSysParam^.astStUnitParam_UnSave[iAxisId].xAxisAlarm_PrnRoller OR i_pstStSysParam^.astStUnitParam_UnSave[iAxisId].xPosDeviationAlarm_PrnRoller);(*轴报警|*)
				pstStIOMap_AxisBasic^.o_xLamp_Inch:= i_pstStSysParam^.astStUnitParam_UnSave[iAxisId].xAxisInching OR g_axAxisInchDecing[iAxisId];(*单运行|*)

 			END_IF
		END_FOR

		//2026.03.26.105424 | + | 挪出来
		//2026.05.20.185157 指针未挪出来 wxy
		pstStIOMap_Main_If:=ADR(i_pastStIOMap_Main^[i_iAxisId_If]);(*读取牵引轴IO|*)
		pstStIOMap_Main_Of:=ADR(i_pastStIOMap_Main^[i_iAxisId_Of]);(*读取牵引轴IO|*)
		IF (i_pstStSysParam^.astStGrpParam_UnSave[i_iGrpId].xFlag_Print AND NOT i_pstStSysParam^.astStGrpParam_UnSave[i_iGrpId].xFlag_FilmAccDecDone) OR
			(i_pstStSysParam^.astStGrpParam_UnSave[i_iGrpId].xFlag_TensionUnfinished) THEN(*张力投入未完成的时候印刷灯闪烁指示@2022.11.30.093228*)
			IF (tmNow-tmLastStateChanged_print)>=T#500ms THEN (* 2021.3.3.114446/改为time()计时方法 *)
				pstStIOMap_Main_If^.o_xLamp_Print:= NOT pstStIOMap_Main_If^.o_xLamp_Print;
				pstStIOMap_Main_Of^.o_xLamp_Print:= NOT pstStIOMap_Main_Of^.o_xLamp_Print;
				//IF iN=1(*i_iGrpAxisNum_PU*) THEN(*检查到最后一个轴更新时间*)
					tmLastStateChanged_print:= tmNow; (* 2021.3.3.114723/ *)
				//END_IF
			END_IF

		ELSE
			pstStIOMap_Main_If^.o_xLamp_Print:=i_pstStSysParam^.astStGrpParam_UnSave[i_iGrpId].xFlag_Print;
			pstStIOMap_Main_Of^.o_xLamp_Print:=i_pstStSysParam^.astStGrpParam_UnSave[i_iGrpId].xFlag_Print;
			tmLastStateChanged_print:= tmNow; (* 2021.3.3.114723/ *)
		END_IF

		IF (i_pstStSysParam^.astStGrpParam_UnSave[i_iGrpId].xFlag_Accing OR i_pstStSysParam^.astStGrpParam_UnSave[i_iGrpId].xFlag_Decing) OR (* 速度在变化中 *)
			i_pstStSysParam^.astStGrpParam_UnSave[i_iGrpId].xFlag_KeepAlarming THEN(*开机响铃的时候闪烁|2022.5.27.123851*)
// 			IF ((i_pstStSysParam^.astStUnitParam_Save[iAxisId].xLinkage AND iN<=i_iGrpAxisNum_PU) OR (* 联动 |只检查色组轴*)
// 				(iN>i_iGrpAxisNum_PU)) THEN(*牵引轴直接处理*)
				IF (tmNow-tmLastStateChanged_prestart)>=T#500ms THEN (* 2021.3.3.114446/改为time()计时方法 *)
					pstStIOMap_Main_If^.o_xLamp_Prestart:= NOT pstStIOMap_Main_If^.o_xLamp_Prestart; (* 2021.3.3.114238/翻转状态 *)
					pstStIOMap_Main_Of^.o_xLamp_Prestart:= NOT pstStIOMap_Main_Of^.o_xLamp_Prestart;
					//IF iN=1(*i_iGrpAxisNum_PU*) THEN(*检查到最后一个轴更新时间*)
						tmLastStateChanged_prestart:= tmNow; (* 记录下这次状态变化的时间 *)
					//END_IF
				END_IF

				(*2021.7.23.144216 altma处理在空转时候闪烁空转灯|印刷时候闪烁印刷灯*)
				IF i_iCustomerNameId=CUSTOMERNAME_ALTMA THEN
					pstStIOMap_Main_If^.o_xLamp_Ink:=pstStIOMap_Main_If^.o_xLamp_Prestart AND i_pstStSysParam^.astStGrpParam_UnSave[i_iGrpId].xFlag_Ink;
					pstStIOMap_Main_If^.o_xLamp_Print:=pstStIOMap_Main_If^.o_xLamp_Prestart AND i_pstStSysParam^.astStGrpParam_UnSave[i_iGrpId].xFlag_Print;
					pstStIOMap_Main_Of^.o_xLamp_Ink:=pstStIOMap_Main_Of^.o_xLamp_Prestart AND i_pstStSysParam^.astStGrpParam_UnSave[i_iGrpId].xFlag_Ink;
					pstStIOMap_Main_Of^.o_xLamp_Print:=pstStIOMap_Main_Of^.o_xLamp_Prestart AND i_pstStSysParam^.astStGrpParam_UnSave[i_iGrpId].xFlag_Print;
				END_IF
			//END_IF
		ELSE
			pstStIOMap_Main_If^.o_xLamp_Prestart:= i_pstStSysParam^.astStGrpParam_UnSave[i_iGrpId].xFlag_PreStart OR i_pstStSysParam^.astStGrpParam_UnSave[i_iGrpId].xFlag_Ink OR i_pstStSysParam^.astStGrpParam_UnSave[i_iGrpId].xFlag_Print;
			pstStIOMap_Main_Of^.o_xLamp_Prestart:= i_pstStSysParam^.astStGrpParam_UnSave[i_iGrpId].xFlag_PreStart OR i_pstStSysParam^.astStGrpParam_UnSave[i_iGrpId].xFlag_Ink OR i_pstStSysParam^.astStGrpParam_UnSave[i_iGrpId].xFlag_Print;
			tmLastStateChanged_prestart:= tmNow; (* 2021.3.3.113954/ *)
		END_IF

		(*收牵指示灯处理|*)
		IF i_iAxisId_Of>=1 AND i_iAxisId_Of<=MAX_UNIT_NUM THEN
			pstStIOMap_Main:= ADR(i_pastStIOMap_Main^[i_iAxisId_Of]);
					pstStIOMap_Main^.o_xLamp_Estop:= i_pstStSysParam^.astStGrpParam_UnSave[i_iGrpId].xFlag_Estop;
					pstStIOMap_Main^.o_xLamp_Stop:= xLamp_Stop;
					pstStIOMap_Main^.o_xLamp_Ink:= i_pstStSysParam^.astStGrpParam_UnSave[i_iGrpId].xFlag_Ink;
					pstStIOMap_Main^.o_xLamp_Tension:= i_pstStSysParam^.astStGrpParam_UnSave[i_iGrpId].xFlag_Tension;
					pstStIOMap_Main^.o_xLamp_AllPress:= i_pstStSysParam^.astStGrpParam_UnSave[i_iGrpId].xFlag_AllPress;(*全体合压灯*)

		END_IF
		(*放牵指示灯处理|*)
		IF i_iAxisId_If>=1 AND i_iAxisId_If<=MAX_UNIT_NUM THEN
			pstStIOMap_Main:= ADR(i_pastStIOMap_Main^[i_iAxisId_If]);
					pstStIOMap_Main^.o_xLamp_Estop:= i_pstStSysParam^.astStGrpParam_UnSave[i_iGrpId].xFlag_Estop;
					pstStIOMap_Main^.o_xLamp_Stop:= xLamp_Stop;
					pstStIOMap_Main^.o_xLamp_Ink:= i_pstStSysParam^.astStGrpParam_UnSave[i_iGrpId].xFlag_Ink;
					pstStIOMap_Main^.o_xLamp_Tension:= i_pstStSysParam^.astStGrpParam_UnSave[i_iGrpId].xFlag_Tension;
					pstStIOMap_Main^.o_xLamp_AllPress:= i_pstStSysParam^.astStGrpParam_UnSave[i_iGrpId].xFlag_AllPress;(*全体合压灯*)

		END_IF

	ELSE
		o_iErNo:= -1;
	END_IF
END_IF

(* ---- KS_FB_GrpUserActionCtrl.st ---- *)
(*@CES
Name=KS_FB_GrpUserActionCtrl
Type=FunctionBlock
TypeGuid=6f9dac99-8de1-4efc-8465-68ac443b7d08
Guid=28236d52-8909-437b-95a9-a6f46f9e83ee
HasDeclaration=True
HasImplementation=True
*)
{DECLARATION}
FUNCTION_BLOCK KS_FB_GrpUserActionCtrl
VAR_INPUT
	i_xEn:BOOL;
	i_iGrpId								: INT;
	i_iCustomerName							: INT;
	i_pastStIOMap_Main_FE					: POINTER TO ARRAY [1..4] OF StIOMap_Main_FE;(*轴io数据区域|*)
	i_pastStIOMap_Axis_FE					: POINTER TO ARRAY [1..MAX_UNIT_NUM] OF StIOMap_Axis_FE;(*轴io数据区域|`````````````````````````````````````````````*)
	i_pastStIOMap_Axis_Extra_FE				: POINTER TO ARRAY [1..MAX_UNIT_NUM] OF StIOMap_Axis_Extra_FE;
	i_pstStIOMap_UwRw_FE_Uw					: POINTER TO ARRAY [1..2] OF StIOMap_UwRw_FE;(*轴io数据区域|*)
	i_pstStIOMap_UwRw_FE_Rw					: POINTER TO ARRAY [1..2] OF StIOMap_UwRw_FE;(*轴io数据区域|*)
	i_iIOGrpIdx_Uw: INT := 1;(*放料组id|*)
	i_iIOGrpIdx_Rw: INT := 1;(*收料组id|*)
	i_iAxisId_If			: INT 						:= -1;(*放牵轴id|*)
	i_iAxisId_Of			: INT 						:= -1;(*收牵轴id|*)
	i_pstStEvtReq: POINTER TO StEvtReq;(*按钮输入操作及边沿触发描述|*)
	i_xInverterAlarm: BOOL;
	i_xBrakeFilm:BOOL;
	i_xLostPressure							: BOOL;(*气压低报警|不允许开机*)
	i_xPrnRollerLoose_AtLeast1				: BOOL;(*至少一色夹板松报警|不允许开机*)
	i_xNeedEstop_BrakeAlarm					: BOOL;(*制动电阻报警急停|2022.5.11.112758*)
	i_paxCommVel_Sure: POINTER TO ARRAY [1..2,1..3] OF BOOL;(*2019.10.21.095108|常用速度123按钮*)
	i_xFalg_ExhaustEn: BOOL;
	i_prVel_Tar_HMI: POINTER TO REAL;
	i_pxTapPosition_Breaking		: POINTER TO BOOL;
	i_pxTapPosition_Printing		: POINTER TO BOOL;
	i_pxTapPosition_UniformInk		: POINTER TO BOOL;
	i_pxAutoAccDec_Hmi				: POINTER TO BOOL;
	i_arVel_CommonlyUsed			: ARRAY [1..3] OF REAL;
	i_xFalg_ExhaustLimitStart: BOOL;
	i_rVel_Cur					: REAL;
	i_rVel_Ink					: REAL;(*空运转速度*)
	i_xFlag_TensionDone:BOOL;
	i_xFlag_TensionUnfinished:BOOL;
	i_xFlag_LinkageAxisAlarm:BOOL;
	i_uiMaxVel_UseCalcAcc: UINT;
	i_pxFlag_KeepAlarming: POINTER TO BOOL;
	i_iTime_Stop: INT;
	i_iTime_FastStop: INT;
	i_iTime_Estop: INT;
	i_iTime_AutoAcc: INT;
	i_iTime_AutoDec: INT;
	i_iTime_ManuAcc: INT;
	i_iTime_ManuDec: INT;
	i_xFilmAccDecDone: BOOL;
	i_byAutoAccDecCurve: BYTE;
	i_iTime_S:INT;
	i_iTime_S_End: INT;
	i_rVel_Max: REAL;
	i_prAccDecTime_ThisTime: POINTER TO REAL;
	i_rAux_enc_vel: REAL;
//	i_pxFlag_FilmAccDecDone							: POINTER TO BOOL; (* 料膜加速完成标志 *)
//	i_uiMaxVel_UseCalcAcc: uint;
	i_xUseMaxTimeAsSBegin_InLowSpeed: BOOL;
	i_rSpeed_SCoeff_Type789: REAL;

END_VAR
VAR_OUTPUT
	o_xEn: BOOL;
	o_iErNo: INT;
	o_xSpeedHigh: BOOL;(*2019.6.14.094543|niu.j|输出速度过高不允许印刷*)
	o_byActionCtlWay: BYTE;(*动作流程选择
							|0:预启动--空转--张力投入--印刷--空转--停机
							|1:预启动--空转--停机;预启动--张力投入--印刷(速度为0)--停机*)
	o_xFlag_FastStoppBtnDn: BOOL;(*2022.4.13.154907 快停被按下了*)
	o_xTips_ExhausLimitStart: BOOL;(*2022.5.21.102417*)
	(*2022.6.28.151929*)
	o_xTowerInvAlarm_Uw					: BOOL;
	o_xTowerInvAlarm_Rw					: BOOL;

	o_iIdGSE								: INT;(*状态!*)
	o_xFlag_Stop							: BOOL;(*停机标志*)
	o_xFlag_PreStart						: BOOL;(*预启动标志|从停机状态按(预)启动置位标志 色组速度达到空转速度清o_xFlag_PreStart标志,置位o_xFlag_Ink标志;当o_xFlag_Print标志有效后,*)
	o_xFlag_PreStart_Print					: BOOL;(*印刷预启动标志|用于华丰逻辑变量*)
	o_xFlag_Ink								: BOOL;(*匀墨标志|>20m/min不能联动*)
	o_xFlag_InkAccing						: BOOL;(*匀墨加速中<指0~10m/min那个加速过程>*)
	o_xFlag_Tension							: BOOL;(*张力投入标志|张力投入有效时收放料变频开始起作用|收放料就位后按印刷按钮,牵引压辊合压|o_xFlag_Print有效时张力投入不处理*)
	o_xFlag_Print							: BOOL;(*张力拉料标志有效时，按联动或印刷按钮 先压收牵(延时2s)再压放牵 印刷标志|印刷色组根据联动标志按用户指定的压辊顺序逐一延时压胶辊|胶辊压合完毕后才可置该标志有效|*)
	o_xFlag_Estop							: BOOL;(*急停标志|和停机一样要减速到0，只不过减速时间是急停时间*)
	o_xFlag_AutoAcc							: BOOL;(*自动加速*)
	o_xFlag_AutoDec							: BOOL;(*自动减速*)
	o_xFlag_ManuAcc							: BOOL;(*手动加速*)
	o_xFlag_ManuDec							: BOOL;(*手动减速*)
	o_xFlag_Accing							: BOOL;(*加速中*)
	o_xFlag_Decing							: BOOL;(*减速中*)
	o_xFlag_EStoping						: BOOL;(*正在急停中*)
	o_xFlag_Stoping							: BOOL;(*停机中*)
	o_xFlag_FastStoping						: BOOL;(*快速停机中*)
	o_xLinkage_IfOf_Ink						: BOOL;
	(*o_xFlag_GotoInking						: BOOL;(*转到匀墨*)*)
	o_xTensionNotFinish						: BOOL;(*按下印刷按钮张力投入未完成输出*)
	o_xToPrintVelTooHigh					: BOOL;(*进入印刷状态时速度太高了*)
	o_rFinalVelocity						: REAL;(*目标速度*)
	o_iTimeSec_AccDec_AllTheWay				: INT;(*全程加减速所需要的秒|*)
	(*2025.2.10.110905+ 单位修改了0.1s@急停的时候需要更短*)
	o_iTimeSec_AccDec_AllTheWay_0_1s		: INT;(*输出时间单位为0.1s*)
	o_xVel_Tar_OverRange					: BOOL;(*目标速度超限值|2019.10.28.102337*)
	o_xFlag_ArrivedToTargetVel				: BOOL;
	o_diVel_Virtual_Tar: dINT;
	o_lrMax_a_S_pos: LREAL;
	o_lrTime_S : LREAL;
	o_lrJerk_SBegin: LREAL;
	o_lrJerk_SEnd: LREAL;
//	o_rVel_Film: REAL;
	o_rVel_PrnRoller								: REAL;(* 版辊运行速度*)
	o_rVel_NetRoller								: REAL;(* 网辊运行速度*)
	o_rVel_BottomRoller								: REAL;(* 底辊运行速度*)
	o_rVel_Cur_HMI									: REAL;(* 当前屏显速度 *)
END_VAR
VAR
	xBtnInk: BOOL;(*空转*)
	xBtnPrint: BOOL;(*印刷*)
	xBtnTension: BOOL;(*张力投入*)
	xBtnManuAcc: BOOL;(*手动加速*)
	xBtnManuDec: BOOL;(*手动减速*)
	xBtnAutoAccOrDec: BOOL;(*自动加减速*)
	xBtnStop: BOOL;(*停止*)
	xBtnFastStop: BOOL;(*快速停止|2022.4.9.235219*)
	xBtnEstop: BOOL;(*急停*)
	lrVel_Tar: LREAL;
	axNeedRstTrig_AutoAccOrDec: ARRAY [1..3] OF BOOL;
	xLastFlag_Stop: BOOL;
	xLastFlag_Ink: BOOL;
	xLastFlag_TensionUnFinished: BOOL;(*2022.11.30.093132*)
	bySpecialProcess:BYTE:=0;(*2022.5.29.001333*)
	tmHold_PreStart: TIME := T#3S; (* 开机预启动持续时间| 2022.5.27.143829*)
	byStates: BYTE;(*2023.09.21.143746 增加*)
	fbTon_Timming: TON;(*2023.12.16.155301*)
	fbKS_FB_StdActionCtl: KS_FB_StdActionCtl;
(*	fbKS_FB_SpeedControl: KS_FB_SpeedControl_2;	*)
	fbKS_FB_SpeedControl_V2: KS_FB_SpeedControl_V2;

(*	fbKS_FB_FilmSpdCtrl: KS_FB_FilmSpdCtrl;*)
	lrServoMotorRatedVel: LREAL;(*伺服电机额定转速可以达到的线速度|*)
	axFlag_PreStart: ARRAY [1..2] OF BOOL;
	xReCalc_Target: BOOL;
	xVel_Tar_OverRange: BOOL;
	xChangeSts_To_Ink: BOOL;
	xChangeSts_To_Prn: BOOL;
END_VAR
VAR_IN_OUT
	io_xMotionEnabled: BOOL;(*|2021.1.15.092801 速度控制块使能修改为输入输出变量|这里处理该值的复位*)
END_VAR
{IMPLEMENTATION}
o_xEn:= i_xEn;
o_iErNo:= 0;
IF i_xEn THEN
	(*1.限速处理稍后再算*)

	(*2.先处理按钮动作*)
	KS_ActionBtnDeal(
		i_iGrpId,(*i_iGrpId,*)
		i_pstStEvtReq,(*i_pstStEvtReq:= , *)
		ADR(o_byActionCtlWay),(*i_pbyActionCtlWay:= , *)
		ADR(xBtnInk),(*i_pxBtnInk:= ,*)
		ADR(xBtnPrint),(*i_pxBtnPrint:= ,*)
		ADR(xBtnTension),(*i_pxBtnTension:= ,*)
		ADR(xBtnManuAcc),(*i_pxBtnManuAcc:= ,*)
		ADR(xBtnManuDec),(*i_pxBtnManuDec:= ,*)
		ADR(xBtnAutoAccOrDec),(*i_pxBtnAutoAccOrDec:= ,*)
		ADR(xBtnStop),(*i_pxBtnStop:= ,*)
		ADR(xBtnFastStop),(*i_pxBtnFastStop:= ,*)
		ADR(xBtnEstop),(*i_pxBtnEstop:= ,*)
		ADR(lrVel_Tar),(*i_plrVel_Tar:= ,*)
		i_xInverterAlarm,(*i_xInverterAlarm:= ,*)
		i_xBrakeFilm,(*i_xBrakeFilm:= ,*)
		i_xLostPressure,(*i_xLostPressure:= ,*)
		i_xPrnRollerLoose_AtLeast1,(*i_xPrnRollerLoose_AtLeast1:= ,*)
		i_xNeedEstop_BrakeAlarm,(*i_xNeedEstop_BrakeAlarm:= ,*)
		i_paxCommVel_Sure,(*i_paxCommVel_Sure:= ,*)
		ADR(axNeedRstTrig_AutoAccOrDec),(*i_paxNeedRstTrig_AutoAccOrDec:= ,*)
		ADR(xLastFlag_Stop),(*i_pxLastFlag_Stop:= ,*)
		ADR(xLastFlag_Ink),(*i_pxLastFlag_Ink:= ,*)
		ADR(xLastFlag_TensionUnFinished),(*i_pxLastFlag_TensionUnFinished:= ,*)
		i_xFalg_ExhaustEn,(*i_xFalg_ExhaustEn:= ,*)
		ADR(o_xFlag_FastStoppBtnDn),(*i_pxFastStopBtnDn:= ,*)
		ADR(o_xTips_ExhausLimitStart),(*i_pxTips_ExhausLimitStart:= ,*)
		ADR(bySpecialProcess),(*i_pbySpecialProcess:= ,*)
		ADR(tmHold_PreStart),(*i_ptmHold_PreStart:= ,*)
		gc_tmHold_PreStart_BeiRen,(*i_tmHold_PreStart_BeiRen:= ,*)
		gc_tmAlarmHold_PreStart,(*i_tmAlarmHold_PreStart:= ,*)
		ADR(byStates),(*i_pbyStates:= ,*)
		ADR(fbTon_Timming),(*i_pfbTon:= ,*)
		i_iCustomerName,(*i_iCustomerName:= ,*)
		ADR(o_xLinkage_IfOf_Ink),(*i_pxLinkage_IfOf_Ink:= ,*)
		i_prVel_Tar_HMI,(*i_prVel_Tar_HMI:= ,*)
		i_pxTapPosition_Breaking ,
		i_pxTapPosition_Printing ,
		i_pxTapPosition_UniformInk,
		i_pxAutoAccDec_Hmi,
		i_arVel_CommonlyUsed,
		i_xFalg_ExhaustLimitStart,
		i_rVel_Ink,(*i_rVel_Ink:= ,*)
		o_xFlag_Stop,(*i_xFlag_Stop:= , *)
		o_xFlag_Estop,(*i_xFlag_Estop:= ,*)
		o_xFlag_Ink,(*i_xFlag_Ink:= ,*)
		o_xFlag_Print,(*i_xFlag_Print:= ,*)
		o_xFlag_InkAccing,(*i_xFlag_InkAccing:= ,*)
		o_xFlag_Stoping,(*i_xFlag_Stoping:= ,*)
		o_xFlag_EStoping,(*i_xFlag_EStoping:= ,*)
		o_xFlag_Tension,(*i_xFlag_Tension:= ,*)
		i_xFlag_TensionDone,
		i_xFlag_TensionUnfinished,
		i_xFlag_LinkageAxisAlarm,
		i_rVel_Cur,(*i_rVel_Cur:= ,*)
		o_xFlag_AutoAcc,(*i_xFlag_AutoDec:= ,*)
		o_xFlag_AutoDec,(*i_xFlag_AutoAcc:= ,*)
		o_xFlag_Accing,(*i_xFlag_Accing:= ,*)
		o_xFlag_Decing,(*i_xFlag_Decing:= *)
		io_xMotionEnabled,
		ADR(xChangeSts_To_Ink),
		ADR(xChangeSts_To_Prn));

	fbKS_FB_StdActionCtl(
		i_xEn:= TRUE,
		i_byActionCtlWay:= o_byActionCtlWay,
		i_xBtnInk:= xBtnInk,
		i_xBtnPrint:= xBtnPrint ,
		i_xBtnTension:= xBtnTension,
		i_xBtnManuAcc:= xBtnManuAcc ,
		i_xBtnManuDec:= xBtnManuDec ,
		i_xBtnAutoAccOrDec:=  xBtnAutoAccOrDec,
		i_xBtnStop:=  xBtnStop,
		i_xBtnFastStop:=  xBtnFaststop,
		i_xBtnEstop:=  xBtnEstop,

		i_xTensionDne:= i_xFlag_TensionDone,
		i_lrVel_Cur:= i_rVel_Cur,
		i_lrVel_Max:= i_rVel_Max,//lrServoMotorRatedVel,		//bai.zy | TEST_ 临时使用 |此处应该是电机最高转速对应的最大速度lrServoMotorRatedVel,
		i_lrVel_Tar:= lrVel_Tar(*i_pstStGrpParam^.lrVel_Tar*) ,
		i_lrVel_Ink:= i_rVel_Ink,
		i_iTime_Ink:= UINT_TO_INT(i_uiMaxVel_UseCalcAcc/5),(*2024.04.12.173848 空转加速时间*)
		i_iTime_Stop:= i_iTime_Stop,
		i_iTime_FastStop:= i_iTime_FastStop,
		(*2025.2.8.162629*)
		i_iTime_Estop:= i_iTime_Estop,
		i_iTime_AutoAcc:= i_iTime_AutoAcc,
		i_iTime_AutoDec:= i_iTime_AutoDec,
		i_iTime_ManuAcc:= i_iTime_ManuAcc,
		i_iTime_ManuDec:= i_iTime_ManuDec,
		i_pxFlag_ArrivedToTargetVel:= ADR(o_xFlag_ArrivedToTargetVel),
		i_pxFlag_KeepAlarming:= i_pxFlag_KeepAlarming,
		i_xFilmAccFinish:= i_xFilmAccDecDone,(*2019.10.08.104841|niu.j|新增料膜加速完成标志*)
		(*2022.5.29.000637*)
		i_tmHold_PreStart:=tmHold_PreStart, (* 开机预启动持续时间| 2022.5.27.143829*)
		i_bySpecialProcess:=bySpecialProcess,(*在基础的开机流程上增加了特殊开机方式切换标志|0:按照基础的|
																						   |1:北人的*)
		i_xBtnInk_BeiRen:=i_pstStEvtReq^.xEvt_Ink,(*空转按钮-专为北人使用|和基础流程的空转按钮定义不同|2022.5.28.234758*)
		i_xEstopTimeIsActTime:=FALSE,(*2025.2.8.163238 不做切换了,就直接修改为输入时间是实际急停时间*)
		i_uiMaxVel_UseCalcAcc:=i_uiMaxVel_UseCalcAcc,
		i_xEstopTimeIsToMaxVel:=TRUE,(*2025.2.13.131137  急停时间是到达最大速度的时间*)
		o_xEn=> ,
		o_iIdGSE=>o_iIdGSE ,
		o_xFlag_Stop=> o_xFlag_Stop,
		o_xFlag_PreStart=> axFlag_PreStart[1],
		o_xFlag_PreStart_Print=> axFlag_PreStart[2],
		o_xFlag_Ink=> o_xFlag_Ink,
		o_xFlag_InkAccing=> o_xFlag_InkAccing,
		o_xFlag_Tension=> o_xFlag_Tension,
		o_xFlag_Print=> o_xFlag_Print,
		o_xFlag_Estop=> o_xFlag_Estop,
		o_xFlag_AutoAcc=> o_xFlag_AutoAcc,
		o_xFlag_AutoDec=> o_xFlag_AutoDec,
		o_xFlag_ManuAcc=> o_xFlag_ManuAcc,
		o_xFlag_ManuDec=> o_xFlag_ManuDec,
		o_xFlag_Accing=> o_xFlag_Accing,
		o_xFlag_Decing=> o_xFlag_Decing,
		o_xFlag_EStoping=> o_xFlag_EStoping,
		o_xFlag_Stoping=> o_xFlag_Stoping,
		o_xFlag_FastStoping=> o_xFlag_FastStoping,
(*			o_xFlag_GotoInking=> i_pstStGrpParam^.xFlag_GotoInking,*)
		o_xTensionNotFinish=> o_xTensionNotFinish,
		o_xReCalc_Target=> xReCalc_Target,
		o_xToPrintVelTooHigh=>o_xSpeedHigh,
		o_rFinalVelocity=> o_rFinalVelocity,
		o_iTimeSec_AccDec_AllTheWay=>,
		(*2025.2.10.113946 按照0.1s单位输出*)
		o_iTimeSec_AccDec_AllTheWay_0_1s=>o_iTimeSec_AccDec_AllTheWay_0_1s,
		o_xVel_Tar_OverRange=>xVel_Tar_OverRange );
	(*速度功能块处理*)
		o_xFlag_PreStart_Print:= axFlag_PreStart[2];
	IF i_iTime_S= 0 THEN
		i_iTime_S:= 30;
	END_IF
	IF i_iTime_S_End=0 THEN
		i_iTime_S_End:=30;
	END_IF
fbKS_FB_SpeedControl_V2(
		i_xEn:= io_xMotionEnabled,
		i_byAutoAccDecCurve:= i_byAutoAccDecCurve,
		i_iMsCycle_Motion:= gc_EXT_TSK_CYCLE_TIME,
		i_lrTimeSec_SBegin:= INT_TO_LREAL(i_iTime_S),
		i_lrTimeSec_SEnd:= INT_TO_LREAL(i_iTime_S_End),
		i_xReCalc_Target:= xReCalc_Target,
		i_piTimeSec_AccDec_AllTheWay:= ADR(o_iTimeSec_AccDec_AllTheWay_0_1s),
		i_rVel_Max:= i_rVel_Max,
		i_pxFlag_ArrivedToTargetVel:= ADR(o_xFlag_ArrivedToTargetVel),
		i_rFinalVelocity:= LREAL_TO_REAL(o_rFinalVelocity),
		i_prVel_Cur:= ADR(i_rVel_Cur),
		i_prAccDecTime_ThisTime:= i_prAccDecTime_ThisTime,
		i_xFlag_PTfifofull:= FALSE,
		i_xFlag_ManuAcc:= o_xFlag_ManuAcc,
		i_xFlag_ManuDec:= o_xFlag_ManuDec,
		i_xFlag_EStoping:= o_xFlag_EStoping,
		i_xFlag_Stoping:= o_xFlag_Stoping,
		i_pxFlag_Decing:= ADR(o_xFlag_Decing),
		i_pxFlag_Accing:= ADR(o_xFlag_Accing),
		i_xFlag_AutoAcc:= o_xFlag_AutoAcc,
		i_xFlag_AutoDec:= o_xFlag_AutoDec,
		i_xFlag_InkAccing:= o_xFlag_InkAccing,
		i_iIdGSE:= o_iIdGSE,
		i_xFlag_Print:= o_xFlag_Print,
		i_xFlag_FastStoping:= o_xFlag_FastStoping,
		i_xFlag_Ink:= o_xFlag_Ink,
		i_rAux_enc_vel:= i_rAux_enc_vel,
		i_rGirth_Master:= gc_rGirth_Master,
		i_uiMaxVel_UseCalcAcc:= i_uiMaxVel_UseCalcAcc,
		i_rSpeed_SCoeff_Type789:= i_rSpeed_SCoeff_Type789,
		i_xUseMaxTimeAsSBegin_InLowSpeed:= i_xUseMaxTimeAsSBegin_InLowSpeed,
		i_iTime_AutoAcc:= i_iTime_AutoAcc,
		i_iTime_AutoDec:= i_iTime_AutoDec,
		o_xEno=> ,
		o_iErNo=> ,
		o_diVel_Virtual_Tar=> o_diVel_Virtual_Tar,
		o_lrMax_a_S_pos=> o_lrMax_a_S_pos,
		o_lrTime_S=> o_lrTime_S,
		o_lrJerk_SBegin=> o_lrJerk_SBegin,
		o_lrJerk_SEnd=> o_lrJerk_SEnd
	);
(*
	fbKS_FB_SpeedControl(
		i_xEn:= io_xMotionEnabled,
		i_byAutoAccDecCurve:= i_byAutoAccDecCurve,
		i_iMsCycle_Motion:= gc_EXT_TSK_CYCLE_TIME,
		i_lrTimeSec_SBegin:= INT_TO_LREAL(i_iTime_S),
		i_lrTimeSec_SEnd:= INT_TO_LREAL(i_iTime_S_End),
		i_xReCalc_Target:= xReCalc_Target,
		i_piTimeSec_AccDec_AllTheWay:= ADR(o_iTimeSec_AccDec_AllTheWay_0_1s),
		i_rVel_Max:= i_rVel_Max,
		i_pxFlag_ArrivedToTargetVel:= ADR(o_xFlag_ArrivedToTargetVel),
		i_rFinalVelocity:= LREAL_TO_REAL(o_lrFinalVelocity),
		i_prVel_Cur:= ADR(i_rVel_Cur),
		i_prAccDecTime_ThisTime:= i_prAccDecTime_ThisTime,
		i_xFlag_PTfifofull:= FALSE,
		i_xFlag_ManuAcc:= o_xFlag_ManuAcc,
		i_xFlag_ManuDec:= o_xFlag_ManuDec,
		i_xFlag_EStoping:= o_xFlag_EStoping,
		i_xFlag_Stoping:= o_xFlag_Stoping,
		i_pxFlag_Decing:= ADR(o_xFlag_Decing),
		i_pxFlag_Accing:= ADR(o_xFlag_Accing),
		i_xFlag_AutoAcc:= o_xFlag_AutoAcc,
		i_xFlag_AutoDec:= o_xFlag_AutoDec,
		i_xFlag_InkAccing:= o_xFlag_InkAccing,
		i_iIdGSE:= o_iIdGSE,
		i_xFlag_Print:= o_xFlag_Print,
		i_xFlag_FastStoping:= o_xFlag_FastStoping,
		i_xFlag_Ink:= o_xFlag_Ink,
		i_rAux_enc_vel:= i_rAux_enc_vel,
		i_rGirth_Master:= gc_rGirth_Master,
		o_xEno=> ,
		o_iErNo=> ,
		o_diVel_Virtual_Tar=> o_diVel_Virtual_Tar,
		o_lrMax_a_S_pos=> o_lrMax_a_S_pos,
		o_lrTime_S => o_lrTime_S);
*)
	//o_rVel_PrnRoller:= o_rVel_Film;//
	//2025.08.07.113103 | bai.zy | TEST_ 临时测试
	o_rVel_PrnRoller:= i_rVel_Cur;
	//o_rVel_BottomRoller:= o_rVel_Film;

	o_rVel_NetRoller:= i_rVel_Cur;
	//o_rVel_BottomRoller:= i_pstStSysParam^.rVel_Film;
	//2025.08.07.113103 | bai.zy | TEST_ 临时测试
	o_rVel_Cur_HMI:= i_rVel_Cur;(* 需要新增 2021.11.6.144801 *)
	//o_rVel_Cur_HMI:= o_rVel_Film;(* 需要新增 2021.11.6.144801 *)

	(*直接调用速度处理|*)
	IF io_xMotionEnabled THEN
		IF (o_xFlag_Stop OR
			o_xFlag_Estop )AND
			i_rVel_Cur=0 THEN
			io_xMotionEnabled:=FALSE;
		END_IF
	END_IF
ELSE
	;
END_IF

(* ---- KS_FB_RollerPressCTL_Home.st ---- *)
(*@CES
Name=KS_FB_RollerPressCTL_Home
Type=FunctionBlock
TypeGuid=6f9dac99-8de1-4efc-8465-68ac443b7d08
Guid=ba8a6c67-74a8-49bb-b69a-0a82809f62f7
HasDeclaration=True
HasImplementation=True
*)
{DECLARATION}
FUNCTION_BLOCK KS_FB_RollerPressCTL_Home
(*2021.10.27.111058 区分联动轴和联动自动合压轴个数*)
(*2022.6.16.134644 增加了放牵延时压辊的参数输入*)
(*2023.2.16.102449兼容张力投入时候收牵合压@牵引手动合压修改了为沿触发了同时收牵离压只处理自动合压的的合压*)
(*2023.07.04.140520 增加接口支持离压到最高点的一些状态处理*)
(*2026.04.10.113911+周期不稳定，延时更换为计时器处理 by liu.yt*)
VAR_INPUT
	i_xEn: BOOL;
	i_iGrpId: INT;
	i_pstStSysParam: POINTER TO StSysParam;
	i_iGrpAxisNum_Pu: INT; (*印刷色组数*)
	i_iAxisId_If: INT;
	i_iAxisId_Of: INT;
	i_pstStEvtReq: POINTER TO StEvtReq;(*按钮输入操作及边沿触发描述|*)
	i_aiGrpAxisList: ARRAY [1..MAX_UNIT_NUM] OF INT; (*系的轴列表|已经按照升序排列了*)
	i_pastStIOMap_Main_FE	: POINTER TO ARRAY [1..4] OF StIOMap_Main_FE;(*轴io数据区域|*)
	i_pastStIOMap_Axis_FE	: POINTER TO ARRAY [1..MAX_UNIT_NUM] OF StIOMap_Axis_FE;(*轴io数据区域|`````````````````````````````````````````````*)
	i_xMachineRev: BOOL;(*反向走料*)
	i_iCycle_Time: INT;
	i_xPressRollerDne_Of_WhenTensionIn:BOOL;(*2023.2.16.112443张力投入时候是否合压收牵标志*)

	(*离压方式-三位五通阀@2023.07.04.140511*)
	i_xUnPressTop_EstopBtn:BOOL;(*急停离压方式标志|FALSE=按照延时离压|TRUE=离压到最高处*)
	i_xUnPressTop_AllUnPressBtn:BOOL;(*全体离压按钮按下时候方式标志|FALSE=按照延时离压|TRUE=离压到最高处*)
	i_xClearUnPressSignal_OnTop:BOOL;(*位于最高点清除离压信号*)
	i_iCycleTime_Plc : INT;
	i_byActionCtlWay: BYTE;(*系动作流程*)
	i_pastStInteraction : POINTER TO ARRAY [1..MAX_UNIT_NUM] OF StInteraction;
END_VAR
VAR_OUTPUT
	o_xEno: BOOL;
	o_xRollerPressDone: BOOL;
END_VAR
VAR

	iCurrentIndex: INT := -1;
	iUnitId: INT;

	iLinkageAxisNum: INT := 0;(*联动轴个数*)
	iAutoPressAxisNum: INT := 0;(*自动压辊轴个数*)
	aiLinkageAxisIdList: ARRAY [1..MAX_UNIT_NUM] OF INT := [MAX_UNIT_NUM(-1)];
	iAutoPressCycleNum: INT;(*自动合压周期计数*)
	iAutoPressNum:INT;(*自动合压的个数*)
	//uiDelayPeriod: UINT:=100;(*抬起压辊延迟的周期数*)
	//周期任务35ms 次数减小一些@2026.04.10.173813+
	uiDelayPeriod: UINT:=50;(*抬起压辊延迟的周期数*)
	iN: INT;
	iCount: INT;
	afbRTrig: ARRAY [1..MAX_UNIT_NUM] OF R_TRIG;
	axPrePress: ARRAY [1..MAX_UNIT_NUM] OF BOOL;

	xInFeed_Press_Delay: BOOL;(*放牵压辊延迟标志有效*)
	iInFeed_Press_DelayNum: INT;(*放牵压辊延时计数*)
	auiFastAdj_UnPressCount: ARRAY [1..MAX_UNIT_NUM] OF INT;
	xAllPress: BOOL;
	xAllUnPress: BOOL;
	fbRTrig_stop1: R_TRIG;
	fbRTrig_stop2: R_TRIG;
	axUnPress_Inching: ARRAY [1..MAX_UNIT_NUM] OF BOOL;	(*点动离压中*)
	xPressDone: BOOL;
	iRollerPressDoneDelay: UINT := 60000;
	xPreStart: BOOL;

	axRel_PressBak: ARRAY [1..MAX_UNIT_NUM] OF BOOL;

	xBtnUnPressTrig: BOOL;(*离压*)
	xUnitPressBtn: BOOL;
	xUnitUnPressBtn: BOOL;

	axPressModeAutoBak:ARRAY [1..MAX_UNIT_NUM] OF BOOL;
	(*2022.5.23.140052*)
	xUnPressForFastStopping: BOOL;(*因为快停需要抬起胶辊*)
	xLastFlag_Sts: BOOL;
	xFlag_FastStoping: BOOL;
	xLastFlag_Tension: BOOL;(*2023.2.16.111933*)
	afbTRIG_Press:ARRAY [1..MAX_UNIT_NUM] OF R_TRIG;
	afbTRIG_UnPress:ARRAY [1..MAX_UNIT_NUM] OF R_TRIG;
	(*2023.07.04.140535*)
	uiTimeMs_RollerPressUpKeep: UINT;
	uiTimeMs_RollerPressUpKeep_OnTop:UINT:=8000;(*离压到最高的时间@MS*)
	abyStsUnPress: ARRAY [1..MAX_UNIT_NUM] OF BYTE;(*离压的状态/=0 离压延时 /=1 离压到最高*)
	byTypeUnPress: BYTE;(*/.0 急停离压到最高/.1 全体离压到最高*)
	fbTrig_TypeUnPress: R_TRIG;
	fbStopToInkTrig: R_TRIG;

(*部分参数需要输入及输出-放这里处理*)
(*输入变量*)
	xFlag_EStoping_In: BOOL;
	xFlag_Estop_In: BOOL;
	xFlag_Print_In: BOOL;
	xFlag_Tension_In: BOOL;
	xFilmAccDecDone_In: BOOL;
	iDelayMsec_RollerPress_In: INT;
	byDelayTime_PressDneInPrint_If_In: BYTE;(*单位是s*)
	xFlag_PreStart_In: BOOL;
	xAllPressOneBtn_In: BOOL;
	xUnitPressOneBtn_In: BOOL;
	xWorkMode_RollerPress_In: BOOL;
	axFlag_Linkage_In: ARRAY [1..MAX_UNIT_NUM] OF BOOL;
	axPressMode_Auto_IO_In: ARRAY [1..MAX_UNIT_NUM] OF BOOL;
	axPressMode_Manu_IO_In: ARRAY [1..MAX_UNIT_NUM] OF BOOL;
	xPressMode_Auto_IO_If_In: BOOL;
	xPressMode_Auto_IO_Of_In: BOOL;
	xPressMode_Manu_IO_If_In: BOOL;
	xPressMode_Manu_IO_Of_In: BOOL;
	axPress_IO_In: ARRAY [1..MAX_UNIT_NUM] OF BOOL;
	axUnPress_IO_In: ARRAY [1..MAX_UNIT_NUM] OF BOOL;
	axUnPress_Inching_In: ARRAY [1..MAX_UNIT_NUM] OF BOOL;
	xTapPosition_Printing_In: BOOL;
	xTapPosition_Breaking_In: BOOL;
	xTapPosition_UniformInk_In: BOOL;
	rVel_Cur_In: REAL;
	rVel_Film_In: REAL;
	xFlag_FastStoping_In: BOOL;
	xFlag_Stop_In: BOOL;
	xFlag_Ink_In: BOOL;
(*输出变量*)
	xFlag_AllPress_Out: BOOL;
	xFlag_AllUnPress_Out: BOOL;
	xRel_Press_IO_If_Out: BOOL;
	xRel_Press_IO_Of_Out: BOOL;

	axRel_Press_IO_Out: ARRAY [1..MAX_UNIT_NUM] OF BOOL;
	axRel_UnPress_IO_Out: ARRAY [1..MAX_UNIT_NUM] OF BOOL;

(*输入输出变量*)
	xFlag_GotoInking_In_Out: BOOL;
	axAxisAutoPressed_In_Out: ARRAY [1..MAX_UNIT_NUM] OF BOOL;
	abyRapidAdjustStep_In_Out: ARRAY [1..MAX_UNIT_NUM] OF BYTE;
//2026.5.14.092403
	abyPrevRapidAdjustStep_Out: ARRAY [1..MAX_UNIT_NUM] OF BYTE;//2026.05.13.204447+ out那里的备份值 by liu.yt

	axRapidAdjust_ing_In_Out: ARRAY [1..MAX_UNIT_NUM] OF BOOL;
	aiRapidAdjust_TimingCnt_In_Out: ARRAY [1..MAX_UNIT_NUM] OF INT;
	auiTimeMs_RollerPressUpKeep_In_Out: ARRAY [1..MAX_UNIT_NUM] OF UINT;
	//2025.9.18.151645+ 手动合压处理初始化@解决旋钮合压按钮再初次上电时压辊合压的问题。
	//必须重新触发才能合压
	xPressBtnDealInit:BOOL;

	//2026.04.10.113935+
	afbUnPressTon:ARRAY [1..MAX_UNIT_NUM] OF TON;//小离压计时器
END_VAR

{IMPLEMENTATION}

(**************************************************************************************
*			压辊控制功能块（色组压辊 以及 收放牵压辊）                                         *
*i_xPressCtrl 为true 时由外部输入压辊信号，false时由输入的按钮控制压辊合压 *
* i_xPositivePress 为 true时从第一色往后压辊，为false时由最后一色色往前压	   *
***************************************************************************************)

IF i_xEn AND
	(i_iGrpId=1 OR i_iGrpId=2) AND
	i_pstStSysParam<>0 AND
	i_iGrpAxisNum_Pu>=1 AND
	i_pastStIOMap_Main_FE<>0 AND
	i_pastStIOMap_Axis_FE<>0 THEN

	Action_Input();

	(*2022.6.16.132522 界面增加牵引压辊延时合压参数*)
	IF i_iCycle_Time<=0 THEN
		i_iCycle_Time:=gc_EXT_TSK_CYCLE_TIME;
	END_IF

	(*2019.08.19.100757|niu.j|预启动抬胶辊*)
	IF xFlag_PreStart_In AND
		xFlag_PreStart_In<>xPreStart THEN
		FOR iN:=1 TO i_iGrpAxisNum_Pu BY 1 DO
			iUnitId:= i_aiGrpAxisList[iN];
			IF axRel_Press_IO_Out[iUnitId] THEN
				axRel_Press_IO_Out[iUnitId]:= FALSE;
				axRel_UnPress_IO_Out[iUnitId]:= TRUE;
			END_IF
		END_FOR
	END_IF
	xPreStart:= xFlag_PreStart_In;

	(*2020.9.8.164916 针对全体合压使用一个按钮还是2个按钮控制进行判断|*)
	IF xAllPressOneBtn_In  THEN(*一个按钮控制*)
		xBtnUnPressTrig:=i_pstStEvtReq^.xReqPressAll;
	ELSE(*两个按钮控制*)
		xBtnUnPressTrig:=i_pstStEvtReq^.xReqUnpressAll;
	END_IF

	IF NOT xFlag_AllPress_Out AND i_pstStEvtReq^.xReqPressAll THEN
		xAllPress:=TRUE;
		xAllUnPress:=FALSE;
(*全体离压处理2023.3.27.103437：||niu*)
	ELSIF (*xFlag_AllPress_Out AND*) xBtnUnPressTrig THEN(*全体离压处理|2023.3.17.103503*)
		xAllPress:=FALSE;
		xAllUnPress:=TRUE;
	ELSE
		xAllPress:=FALSE;
		xAllUnPress:=FALSE;
	END_IF

	iAutoPressAxisNum:= 0;
	iLinkageAxisNum:=0;(*2021.10.27.111037*)
	IF NOT xWorkMode_RollerPress_In THEN(*从后往前顺序压辊|*)
		FOR iN:=i_iGrpAxisNum_Pu TO 1 BY -1 DO
			iUnitId:= i_aiGrpAxisList[iN];
			IF iUnitId>=1 AND iUnitId<=MAX_UNIT_NUM THEN
				IF axFlag_Linkage_In[iUnitId] THEN
					iLinkageAxisNum:=iLinkageAxisNum+1;
					IF  axPressMode_Auto_IO_In[iUnitId] THEN(*2021.10.27.111000*)
						iAutoPressAxisNum:= iAutoPressAxisNum+1;
						aiLinkageAxisIdList[iAutoPressAxisNum]:= i_aiGrpAxisList[iN];
					END_IF
				END_IF
			END_IF
		END_FOR
	ELSE (*顺序压辊*)
		FOR iN:=1 TO i_iGrpAxisNum_Pu BY 1 DO
			iUnitId:= i_aiGrpAxisList[iN];
			IF iUnitId>=1 AND iUnitId<=MAX_UNIT_NUM THEN
				IF axFlag_Linkage_In[iUnitId]  THEN
					iLinkageAxisNum:=iLinkageAxisNum+1;
					IF axPressMode_Auto_IO_In[iUnitId]  THEN
						iAutoPressAxisNum:= iAutoPressAxisNum+1;
						aiLinkageAxisIdList[iAutoPressAxisNum]:= i_aiGrpAxisList[iN];
					END_IF
				END_IF
			END_IF
		END_FOR
	END_IF

(*自动压辊*)

	IF xFlag_Print_In  THEN (*印刷状态才能进行自动压辊*)
		xFlag_GotoInking_In_Out:=TRUE;
		IF NOT  xFlag_AllPress_Out THEN
			IF xAllPress AND xFilmAccDecDone_In  THEN (*自动合压*)
				xFlag_AllPress_Out:=TRUE;
				iAutoPressCycleNum:=0;
			END_IF
		ELSE(*全体合压状态*)
			iAutoPressNum:=0;
			FOR iN:=1 TO iAutoPressAxisNum BY 1 DO
				iUnitId:= aiLinkageAxisIdList[iN];
				IF iUnitId>=1 AND iUnitId<=MAX_UNIT_NUM THEN
					IF NOT axAxisAutoPressed_In_Out[iUnitId] THEN (*自动未合压过*)
						IF NOT axRel_Press_IO_Out[iUnitId] THEN (*未合压*)
							IF iAutoPressNum =0 THEN
								axRel_Press_IO_Out[iUnitId]:=TRUE;
								axRel_UnPress_IO_Out[iUnitId]:=FALSE;
								axAxisAutoPressed_In_Out[iUnitId]:=TRUE;
								iAutoPressNum:=1;
							ELSE
								(*IF iAutoPressCycleNum*i_iCycleTime_Plc>=pstStGrpParam^.iMillisecondsDelay_RollerPress THEN*)
								IF iAutoPressCycleNum*i_iCycleTime_Plc>=iDelayMsec_RollerPress_In THEN
									axRel_Press_IO_Out[iUnitId]:=TRUE;
									axRel_UnPress_IO_Out[iUnitId]:=FALSE;
									axAxisAutoPressed_In_Out[iUnitId]:=TRUE;
									iAutoPressNum:=iAutoPressNum+1;
									iAutoPressCycleNum:=0;
								ELSE
									iAutoPressCycleNum:=iAutoPressCycleNum+1;
									EXIT;
								END_IF
							END_IF
						ELSE(*合压了*)
							axAxisAutoPressed_In_Out[iUnitId]:=TRUE;
							iAutoPressNum:=iAutoPressNum+1;
						END_IF
					ELSE
						(*2020.10.10.111710 取消这段代码|Liu.yt*)
						(*IF NOT  axRel_Press_IO_Out[iUnitId] THEN
							axRel_Press_IO_Out[iUnitId]:=TRUE;
							axRel_UnPress_IO_Out[iUnitId]:=FALSE;
						END_IF*)
						IF NOT axPressModeAutoBak[iUnitId] AND
							axPressMode_Auto_IO_In[iUnitId] THEN(*自动合压完成以后如果
																		手自动旋钮由手动切换到自动时我们合压*)
							axRel_Press_IO_Out[iUnitId]:=TRUE;
							axRel_UnPress_IO_Out[iUnitId]:=FALSE;
						END_IF
						iAutoPressNum:=iAutoPressNum+1;
					END_IF
				END_IF
			END_FOR
		END_IF

		(*更新保存的自动按钮状态变量2020.10.10.112410*)
		FOR iN:=1 TO i_iGrpAxisNum_Pu BY 1 DO
			iUnitId:=i_aiGrpAxisList[iN];
			axPressModeAutoBak[iUnitId]:=axPressMode_Auto_IO_In[iUnitId];(*自动按钮上个周期变量*)
		END_FOR

		(*放牵*)
		IF i_iAxisId_If>=1 AND i_iAxisId_If<=MAX_UNIT_NUM THEN
			IF NOT xRel_Press_IO_If_Out AND(*放牵未合压*)
					xPressMode_Auto_IO_If_In THEN(*放牵在自动状态*)
				IF NOT xInFeed_Press_Delay THEN(*压辊延迟无效*)
					(*2026.06.02.211129 计数单位错误*)
					IF iInFeed_Press_DelayNum * i_iCycle_Time >=byDelayTime_PressDneInPrint_If_In * 1000 THEN
						iInFeed_Press_DelayNum:=0;
						xInFeed_Press_Delay:=TRUE;
					ELSE
						iInFeed_Press_DelayNum:=iInFeed_Press_DelayNum+1;
					END_IF
				END_IF
			END_IF
			IF xInFeed_Press_Delay THEN (*放牵压辊延迟标志有效*)
				xRel_Press_IO_If_Out:= xPressMode_Auto_IO_If_In;
			END_IF
		END_IF
	ELSE(*非印刷状态*)
		xFlag_AllPress_Out:=FALSE;
	END_IF

	(*2023.2.16.112143调整*)
	(*收放牵压辊控制*)
	(*收牵*)
	IF xFlag_Print_In OR
		(xFlag_Tension_In AND i_xPressRollerDne_Of_WhenTensionIn)THEN(*张力投入时收牵压辊*)
		IF i_iAxisId_Of>=1 AND i_iAxisId_Of<=MAX_UNIT_NUM THEN
			xRel_Press_IO_Of_Out:=xPressMode_Auto_IO_Of_In;
		END_IF
	END_IF

(*快速调整时压辊控制*)
	FOR iN:=1 TO i_iGrpAxisNum_Pu BY 1 DO
		iUnitId:= i_aiGrpAxisList[iN];
		IF iUnitId>=1 AND iUnitId<=MAX_UNIT_NUM THEN
  			IF abyRapidAdjustStep_In_Out[iUnitId]=0 THEN
				IF axRapidAdjust_ing_In_Out[iUnitId] THEN (*处于快速调整中状态，说明调整已经结束了*)
					(*取压辊快速对版之前的状态*)
					axRel_Press_IO_Out[iUnitId]:= axRel_PressBak[iUnitId];
					axRel_UnPress_IO_Out[iUnitId]:= NOT axRel_PressBak[iUnitId];
					axRapidAdjust_ing_In_Out[iUnitId]:= FALSE;
					aiRapidAdjust_TimingCnt_In_Out[iUnitId]:=0;

					//2025.12.31.152043 | +
					i_pastStInteraction^[iUnitId].o_xCoarseAdjStart := FALSE;
					i_pastStInteraction^[iUnitId].o_xCoarseAdjEnd := TRUE;
				END_IF
				axRel_PressBak[iUnitId]:=axRel_Press_IO_Out[iUnitId];(*保存调整前的压辊状态*)
			ELSIF abyRapidAdjustStep_In_Out[iUnitId]=1 OR abyRapidAdjustStep_In_Out[iUnitId]=2 THEN
				(*准备进入快速调整状态，等待压辊离压，延迟后进入快速调整状态*)
				IF i_pstStSysParam^.stStSysParam_Save.iCustomerId = CUSTOMERNAME_QINHUA THEN
					axRapidAdjust_ing_In_Out[iUnitId]:= TRUE;
					axRel_UnPress_IO_Out[iUnitId]:= TRUE;
					axRel_Press_IO_Out[iUnitId]:= FALSE;
					IF abyRapidAdjustStep_In_Out[iUnitId]=1 THEN

						//2025.12.31.152043 | +
						i_pastStInteraction^[iUnitId].o_xCoarseAdjStart := TRUE;
						i_pastStInteraction^[iUnitId].o_xCoarseAdjEnd := FALSE;
						IF i_pastStInteraction^[iUnitId].i_xPressRetractionPositionSignal THEN
							abyRapidAdjustStep_In_Out[iUnitId]:=2;
						ELSE
							//2026.1.15.120614 | + | 如果没有信号就超时
							IF aiRapidAdjust_TimingCnt_In_Out[iUnitId]>=uiDelayPeriod THEN
								aiRapidAdjust_TimingCnt_In_Out[iUnitId]:=0;
								abyRapidAdjustStep_In_Out[iUnitId]:=2;
							ELSE
								aiRapidAdjust_TimingCnt_In_Out[iUnitId]:=aiRapidAdjust_TimingCnt_In_Out[iUnitId]+1;
							END_IF
						END_IF
					END_IF
				ELSE
					axRapidAdjust_ing_In_Out[iUnitId]:= TRUE;
					axRel_UnPress_IO_Out[iUnitId]:= TRUE;
					axRel_Press_IO_Out[iUnitId]:= FALSE;
					IF abyRapidAdjustStep_In_Out[iUnitId]=1 THEN
						IF aiRapidAdjust_TimingCnt_In_Out[iUnitId]>=uiDelayPeriod THEN
							aiRapidAdjust_TimingCnt_In_Out[iUnitId]:=0;
							abyRapidAdjustStep_In_Out[iUnitId]:=2;
						ELSE
							aiRapidAdjust_TimingCnt_In_Out[iUnitId]:=aiRapidAdjust_TimingCnt_In_Out[iUnitId]+1;
						END_IF
					END_IF
				END_IF
			ELSE
				abyRapidAdjustStep_In_Out[iUnitId]:=0;
				axRapidAdjust_ing_In_Out[iUnitId]:= FALSE;
				aiRapidAdjust_TimingCnt_In_Out[iUnitId]:=0;
			END_IF
		END_IF
	END_FOR

(*色组压辊手动*)
//2025.9.18.151806+ 手动合压沿处理变量初始化
	IF NOT xPressBtnDealInit THEN
		xPressBtnDealInit:=TRUE;
		FOR iN:=1 TO i_iGrpAxisNum_Pu BY 1 DO
			iUnitId:= i_aiGrpAxisList[iN];
			IF iUnitId>=1 AND iUnitId<=MAX_UNIT_NUM THEN
				//2025.9.18.152157 只处理两个按钮控制形式,应该问题不大！
				afbTRIG_Press[iUnitId](CLK:= axPress_IO_In[iUnitId]);
				afbTRIG_UnPress[iUnitId](CLK:= axUnPress_IO_In[iUnitId]);
			END_IF
		END_FOR
	END_IF
	//end
	IF NOT xFlag_Estop_In THEN (*急停状态不能压辊*)
		FOR iN:=1 TO i_iGrpAxisNum_Pu BY 1 DO
			iUnitId:= i_aiGrpAxisList[iN];
			IF iUnitId>=1 AND iUnitId<=MAX_UNIT_NUM THEN
				(*2020.9.8.170013 色组合压离压按钮单个多个控制选择逻辑|Liu.yt*)
				xUnitPressBtn:=FALSE;
				xUnitUnPressBtn:=FALSE;
				IF xUnitPressOneBtn_In THEN(*单个按钮控制*)
					IF axPress_IO_In[iUnitId] AND
						NOT axPrePress[iUnitId] THEN(*合压按下沿*)
						xUnitPressBtn:=NOT axRel_Press_IO_Out[iUnitId];
						xUnitUnPressBtn:= axRel_Press_IO_Out[iUnitId];
					END_IF
				ELSE(*多个按钮控制*)
					xUnitPressBtn:= axPress_IO_In[iUnitId];
					xUnitUnPressBtn:= axUnPress_IO_In[iUnitId];
				END_IF
				axPrePress[iUnitId]:= axPress_IO_In[iUnitId];
		(*修改为沿触发-2023.3.30.133052适应三档开关*)
				afbTRIG_Press[iUnitId](CLK:= xUnitPressBtn);
				afbTRIG_UnPress[iUnitId](CLK:= xUnitUnPressBtn);
				afbRTrig[iN](CLK:=axPressMode_Manu_IO_In[iUnitId]);(*手动按钮上升沿*)
			(*手动按钮删除手动条件|2020.10.10.110559|Liu.yt*)
			(*	IF  pstStIOMap_AxisBasic^.i_xPressMode_Manu THEN(*手动*)*)
					IF (*xUnitPressBtn*) afbTRIG_Press[iUnitId].Q AND NOT axRel_Press_IO_Out[iUnitId] THEN (*合压*)
						axRel_Press_IO_Out[iUnitId]:= TRUE;
						axRel_UnPress_IO_Out[iUnitId]:= FALSE;
					ELSIF (*xUnitUnPressBtn *) afbTRIG_UnPress[iUnitId].Q AND NOT axRel_UnPress_IO_Out[iUnitId] THEN (*离压*)
						axRel_Press_IO_Out[iUnitId]:= FALSE;
						axRel_UnPress_IO_Out[iUnitId]:= TRUE;
					ELSIF axAxisAutoPressed_In_Out[iUnitId] AND afbRTrig[iN].Q  THEN (*自动合压过*)
						axRel_Press_IO_Out[iUnitId]:= FALSE;
						axRel_UnPress_IO_Out[iUnitId]:= TRUE;
					END_IF
(*					END_IF*)

				(*2018.8.1.104126 |  niu.j | 点动离压*)

				IF  axRel_Press_IO_Out[iUnitId]  THEN
					axRel_UnPress_IO_Out[iUnitId]:= FALSE;
				END_IF
				IF axUnPress_Inching_In[iUnitId] THEN
					(*手动点动离压按钮删除手动条件|2020.10.10.110559|Liu.yt*)
					axUnPress_Inching[iN]:=TRUE;
					(*IF  pstStIOMap_AxisBasic^.i_xPressMode_Manu THEN (*手动状态*)*)
						axRel_UnPress_IO_Out[iUnitId]:= TRUE;
						axRel_Press_IO_Out[iUnitId]:= FALSE;
				(*	ELSIF pstStIOMap_AxisBasic^.i_xPressMode_Auto THEN
						IF NOT pstStGrpParam^.xFlag_AllPress THEN
							pstStIOMap_AxisBasic^.o_xRel_UnPress:= TRUE;
							pstStIOMap_AxisBasic^.o_xRel_Press:= FALSE;
						END_IF
					END_IF*)
				ELSIF axUnPress_Inching[iN] AND NOT axUnPress_Inching_In[iUnitId] THEN
					//axRel_Press_IO_Out[iUnitId]:= FALSE;
					//2026.04.08.165318 变量写错了
					axRel_UnPress_IO_Out[iUnitId]:= FALSE;
					axUnPress_Inching[iN]:=FALSE;
				END_IF

				IF axRel_Press_IO_Out[iUnitId] THEN
					;
				END_IF

			END_IF

		END_FOR
	ELSE;
	END_IF

	IF xPressMode_Manu_IO_If_In THEN
		xRel_Press_IO_If_Out:= TRUE;
	ELSIF xPressMode_Auto_IO_If_In THEN
		;
	ELSE
		xRel_Press_IO_If_Out:= FALSE;
	END_IF
	IF xPressMode_Manu_IO_Of_In THEN
		xRel_Press_IO_Of_Out:= TRUE;
	ELSIF xPressMode_Auto_IO_Of_In THEN
		;
	ELSE
		xRel_Press_IO_Of_Out:= FALSE;
	END_IF
	(*2023.07.04.141713 重新处理了离压方式*)
	(*2023.07.04.140920 移动到此处*)

	byTypeUnPress:=0;
	IF i_xUnPressTop_EstopBtn THEN(*急停离压到最高处*)
		IF	i_pstStEvtReq^.xEvt_Estop OR
			i_pstStEvtReq^.xReqEstop OR
			xFlag_Estop_In OR
			xFlag_EStoping_In THEN
			byTypeUnPress.0:=TRUE;
		END_IF
	END_IF
	IF i_xUnPressTop_AllUnPressBtn THEN(*全体离压按钮离压到最高处@*)
		IF xFlag_AllPress_Out AND xAllUnPress THEN(*按钮按下之后在下面才清除标志呢|放置的位置很重要*)
			byTypeUnPress.1:=TRUE;
		END_IF
	END_IF

	fbTrig_TypeUnPress(CLK:=byTypeUnPress<>0);(*检查是否要离压到最高处沿*)
	FOR iN:=1 TO i_iGrpAxisNum_PU BY 1 DO
		iUnitId:= i_aiGrpAxisList[iN];
		IF iUnitId>=1 AND iUnitId<=MAX_UNIT_NUM THEN
			uiTimeMs_RollerPressUpKeep:= auiTimeMs_RollerPressUpKeep_In_Out[iUnitId];

			(*状态处理*)
			IF axRel_Press_IO_Out[iUnitId] THEN(*合压了就复位成延时离压方式*)
				abyStsUnPress[iUnitId]:=0;
			END_IF
			IF fbTrig_TypeUnPress.Q THEN(*离压到最高点*)
				IF axRel_Press_IO_Out[iUnitId] THEN(*合压的状态切换下*)
					abyStsUnPress[iUnitId]:=1;
				END_IF
			END_IF

			(*延时处理*)
			IF abyStsUnPress[iUnitId]=1 THEN(*离压到最高*)
				IF i_xClearUnPressSignal_OnTop THEN(*在最高点需要清除*)
					uiTimeMs_RollerPressUpKeep:=uiTimeMs_RollerPressUpKeep_OnTop;
				ELSE(*在最高点不需要清除*)
					uiTimeMs_RollerPressUpKeep:=0;
				END_IF
			ELSE(*延时离压*);
(*				uiTimeMs_RollerPressUpKeep;*)
			END_IF
			IF axRel_UnPress_IO_Out[iUnitId] AND NOT axUnPress_Inching_In[iUnitid] THEN
// 				IF uiTimeMs_RollerPressUpKeep<>0 THEN
// 					IF uiTimeMs_RollerPressUpKeep<= i_iCycleTime_Plc*auiFastAdj_UnPressCount[iUnitId] THEN
// 						axRel_UnPress_IO_Out[iUnitId]:= FALSE;
// 					ELSE
// 						auiFastAdj_UnPressCount[iUnitId]:= auiFastAdj_UnPressCount[iUnitId]+1;
// 					END_IF
// 				ELSE
// 					auiFastAdj_UnPressCount[iUnitId]:= 0;
// 				END_IF
				//2026.04.10.114225 重写
				afbUnPressTon[iUnitId](IN:=uiTimeMs_RollerPressUpKeep<>0,PT:=UINT_TO_TIME(uiTimeMs_RollerPressUpKeep));//2026.04.10.114050+
				IF afbUnPressTon[iUnitId].Q THEN//时间到
					axRel_UnPress_IO_Out[iUnitId]:= FALSE;
				END_IF
			ELSE
				auiFastAdj_UnPressCount[iUnitId]:= 0;
				afbUnPressTon[iUnitId](IN:=FALSE);
			END_IF
		END_IF
	END_FOR

	(*条件优化下2023.2.16.112340*)
	IF i_byActionCtlWay=1 THEN(*华丰类似流程@2023.2.16.105907*)
		IF xTapPosition_Printing_In THEN
			fbRTrig_stop1(CLK:=i_pstStEvtReq^.xReqStop AND rVel_Cur_In=0);
			fbRTrig_stop2(CLK:=FALSE);
		ELSIF xTapPosition_Breaking_In OR
			xTapPosition_UniformInk_In THEN
			fbRTrig_stop1(CLK:=FALSE);
			fbRTrig_stop2(CLK:=i_pstStEvtReq^.xReqStop);
		END_IF
	ELSE(*常规流程*);
		fbRTrig_stop1(CLK:=FALSE);
		fbRTrig_stop2(CLK:=FALSE);
	END_IF

	(*2022.5.23.140104*)
	IF xFlag_FastStoping_In THEN
		xFlag_FastStoping:=TRUE;
	END_IF
	xUnPressForFastStopping:=FALSE;
	IF xFlag_FastStoping THEN
		IF xFlag_Stop_In AND
			NOT xLastFlag_Sts THEN(*进入停止状态*)
			xUnPressForFastStopping:=TRUE;
		END_IF

		IF xFlag_Stop_In THEN(*清除标志*)
			xFlag_FastStoping:=FALSE;
		END_IF
	END_IF
	xLastFlag_Sts:= xFlag_Stop_In OR xFlag_EStop_In;
	(*2023.07.04.193801*)
	fbStopToInkTrig(CLK:=xFlag_GotoInking_In_Out  AND xFlag_Ink_In);

(*全体离压处理2023.3.27.103624|niu.*)
	IF ((*pstStGrpParam^.xFlag_AllPress AND*) xAllUnPress) OR(*全体合压状态下 按下了全体离压清除所有压辊输出*)
		fbRTrig_stop1.Q OR
		fbRTrig_stop2.Q OR
		xUnPressForFastStopping OR(*2022.5.23.140354*)
		(*(pstStGrpParam^.xFlag_GotoInking  AND pstStGrpParam^.xFlag_Ink)*)
		fbStopToInkTrig.Q OR (*从印刷状态退出到空转状态@2023.07.04.193731 改成沿触发*)
		xFlag_Estop_In THEN(*急停状态清除压辊输出*)
		FOR iN:=1 TO i_iGrpAxisNum_PU BY 1 DO
			iUnitId:= i_aiGrpAxisList[iN];
			IF iUnitId>=1 AND iUnitId<=MAX_UNIT_NUM THEN
				axRel_Press_IO_Out[iUnitId]:=FALSE;
				axRel_UnPress_IO_Out[iUnitId]:=TRUE;
				axAxisAutoPressed_In_Out[iUnitId]:=FALSE;
(*全体离压处理2023.3.27.103735|niu.*)
				IF NOT ((*pstStGrpParam^.xFlag_AllPress AND*) xAllUnPress) THEN(*全体离压的时候不清除快速对版相关变量*)
					abyRapidAdjustStep_In_Out[iUnitId]:=0;(*清除快速对版相关变量*)
					axRapidAdjust_ing_In_Out[iUnitId]:=FALSE;
					aiRapidAdjust_TimingCnt_In_Out[iUnitId]:=0;

				END_IF
			END_IF
		END_FOR
		(*pstStGrpParam^.xFlag_GotoInking:=FALSE;*)
		xFlag_AllPress_Out:=FALSE;
	END_IF

(*清除收放牵压辊信号*)
	IF (* pstStGrpParam^.lrVel_Film=0 (*AND pstStGrpParam^.iIdGSE<>GSE_PRINT_PRESTART OR
		pstStGrpParam^.xFlag_Stop*) OR*)(*料膜速度=0,并且是从印刷状态停到空转状态*)
		fbRTrig_stop1.Q OR
		fbRTrig_stop2.Q OR
(*2023.2.16.105134屏蔽预启动清除压辊*)
(*		pstStGrpParam^.xFlag_PreStart OR(*预启动时候清除压辊输出*)*)
		(i_xPressRollerDne_Of_WhenTensionIn AND (xLastFlag_Tension AND NOT xFlag_Tension_In))OR(*退出张力投入取消收牵压辊*)
		(xFlag_GotoInking_In_Out AND xFlag_Ink_In(* (rVel_Film_In=0 AND i_byActionCtlWay=0)*)) OR (*从印刷状态退出到空转状态*)
																			(*g_abyActionCtlWay[i_iGrpId]<>2修改为=0|2019.11.28.104528_*)
		xFlag_Estop_In THEN(*急停状态清除压辊输出*)

		IF NOT xPressMode_Manu_IO_If_In THEN(*非手动时清除@2023.2.16.111739*)
			xRel_Press_IO_If_Out:=FALSE;(*清除放牵压辊*)
			xInFeed_Press_Delay:=FALSE;
			iInFeed_Press_DelayNum:=0;
		END_IF

		IF NOT xPressMode_Manu_IO_Of_In THEN(*非手动时清除@2023.2.16.111739*)
			xRel_Press_IO_Of_Out:=FALSE;(*清除收牵压辊*)
		END_IF

		xFlag_GotoInking_In_Out:= FALSE;
	END_IF
	(*2023.2.16.105207*)
	xLastFlag_Tension:= xFlag_Tension_In;

	(*反向走料禁止压辊*)
	FOR iN:=1 TO i_iGrpAxisNum_Pu BY 1 DO
		iUnitId:= i_aiGrpAxisList[iN];
		IF iUnitId>=1 AND iUnitId<=MAX_UNIT_NUM THEN
			IF i_xMachineRev THEN
				IF axRel_Press_IO_Out[iUnitId] THEN
					axRel_Press_IO_Out[iUnitId]:=FALSE;
					axRel_UnPress_IO_Out[iUnitId]:=TRUE;
				END_IF
			END_IF
		END_IF
	END_FOR

	FOR iN:=1 TO i_iGrpAxisNum_Pu BY 1 DO (*判断至少合压一色*)
		iUnitId:= i_aiGrpAxisList[iN];
		IF iUnitId>=1 AND iUnitId<=MAX_UNIT_NUM THEN
			IF axFlag_Linkage_In[iUnitId] THEN
				IF NOT axRel_Press_IO_Out[iUnitId] THEN
					xPressDone:=FALSE;(*至少一色合压*)
				ELSE
					xPressDone:=TRUE;
					EXIT;
				END_IF
			END_IF
		END_IF
	END_FOR

	FOR iN:=1 TO i_iGrpAxisNum_Pu BY 1 DO (*判断全体色组合压完成*)
		iUnitId:= i_aiGrpAxisList[iN];
		IF iUnitId>=1 AND iUnitId<=MAX_UNIT_NUM THEN
			IF axFlag_Linkage_In[iUnitId] THEN
				IF axRel_Press_IO_Out[iUnitId] THEN
					o_xRollerPressDone:=TRUE;
				ELSE
					o_xRollerPressDone:=FALSE;
					EXIT;
				END_IF
			END_IF
		END_IF
	END_FOR
	(*2021.10.27.111121 修改为联动轴个数计时*)
	iRollerPressDoneDelay:= INT_TO_UINT((iLinkageAxisNum+2)*iDelayMsec_RollerPress_In);
	IF NOT o_xRollerPressDone AND xPressDone THEN (*2018.10.6.090512|niu.j*)
		IF iCount< UINT_TO_INT(iRollerPressDoneDelay)/i_iCycle_Time THEN
			iCount:=iCount+1;
		ELSE
			o_xRollerPressDone:= TRUE;
		END_IF
	ELSIF NOT xPressDone THEN
		iCount:=0;
	END_IF

ELSE
	iCurrentIndex:= -1;
END_IF

Action_Output();

(* ---- KS_FB_SpeedControl_2.st ---- *)
(*@CES
Name=KS_FB_SpeedControl_2
Type=FunctionBlock
TypeGuid=6f9dac99-8de1-4efc-8465-68ac443b7d08
Guid=3721ed5a-e7f4-4c95-a3b8-3e53b0c929eb
HasDeclaration=True
HasImplementation=True
*)
{DECLARATION}
FUNCTION_BLOCK KS_FB_SpeedControl_2(*先用这个吧，后面再整理2025.6.12.174817*)
(*变化速度的时候置1次xFlag_ArrivedToTargetVel为TRUE就可以了|*)
(*2022.10.27.164825 修改了第4中速度控制方式未在本次时间基础上前后各加s*)
(*2022.10.27.162617调整|在小于S加减速时间的情况下
						使用本次时间+前后i_bySTime_AtLeast时间的s||2022.12.7.170426*)
(*王宁涛处理了前后s分开问题@2023.3.2.210705*)
(*在空转时候自动加减速修改为了手动方式|Liu.yt@2023.3.2.210734*)
VAR_INPUT
	i_xEn: BOOL;
	i_byAutoAccDecCurve:BYTE;(*2022.4.21.231635|
							默认 按照最大直线加速度进行s处理-
						 	1：按照直线加速时间进行s处理-不限制最大加速度
						 	2：按照直线加速时间进行s处理-限制最大加速度
						 	3：按照直线加速时间全程s处理-
							4: 和默认处理方式接近|使用本次时间+前后i_bySTime_AtLeast时间的s|2022.12.7.170445*)
	i_iMsCycle_Motion: INT;(*运动周期|*)
	i_lrTimeSec_SBegin: LREAL := 30;(*S规划前半程时间|*)
	i_lrTimeSec_SEnd: LREAL := 30;(*S规划后半程时间|*)
	i_xReCalc_Target:BOOL;
	i_piTimeSec_AccDec_AllTheWay					: POINTER TO INT; (* S加减速时间 *)
	i_rVel_Max										: REAL; (* 最大速度 *)
	i_pxFlag_ArrivedToTargetVel						: POINTER TO BOOL; (* | *)
	i_rFinalVelocity								: REAL; (* 加减速末端速度 *)
	i_prVel_Cur										: POINTER TO REAL; (* 当前速度 *)
	i_prAccDecTime_ThisTime							: POINTER TO REAL; (* 本次加减速时间 *)
	i_xFlag_PTfifofull								: BOOL; (* 允许写PT使能 *)
	i_xFlag_ManuAcc									: BOOL; (* 手动加速标志 *)
	i_xFlag_ManuDec									: BOOL; (* 手动减速标志 *)
	i_xFlag_EStoping								: BOOL; (* 急停中标志 *)
	i_xFlag_Stoping									: BOOL; (* 停机中标志 *)
	i_pxFlag_Decing									: POINTER TO BOOL; (* 减速中 *)
	i_pxFlag_Accing									: POINTER TO BOOL; (* 加速中 *)
	i_xFlag_AutoAcc									: BOOL; (* 自动减速 *)
	i_xFlag_AutoDec									: BOOL; (* 自动减速 *)
	i_xFlag_InkAccing								: BOOL; (* 空转加速中 *)
	i_iIdGSE										: INT; (* 当前运行步骤 *)
	i_xFlag_Print									: BOOL;
	i_xFlag_FastStoping								: BOOL;
	i_xFlag_Ink										: BOOL;
	(*i_apstStTravelLogRec: ARRAY [1..GC_LOG_CLASSES_MAX_NUM] OF POINTER TO StTravelLogRec; (* 2021.7.5.144816/ *)*)
(*	i_bySTime_AtLeast:BYTE;(*至少s加减速时间|默认10s*)*)(*需要删除|2023.03.02.112331*)
	i_rAux_enc_vel									: REAL;//虚拟主轴的速度//当速度到位标志触发时，直接将虚拟主轴速度给目标速度
	i_rGirth_Master: REAL;
END_VAR
VAR_OUTPUT
	o_xEno: BOOL;
	o_iErNo: INT;(*0.no error\-1.bad parameters\-2.bad lrVelMax&TimeAccDec|*)
	o_diVel_Virtual_Tar: DINT;
	o_lrMax_a_S_pos: LREAL;
	o_lrTime_S : LREAL;
END_VAR
VAR

	lrVel_delta: LREAL;(*速度变化量|*)
	lrJerk_SBegin: LREAL;
	lrJerk_SEnd: LREAL;
	lrAve_a: LREAL;(*全程平均加速度|*)
	lrMax_a_S: LREAL;(*S规划的最大加速度|*)
	iNum_InflectionPts: INT;
	lrCurr_t: LREAL;(*当前时间|*)
	lrPrev_t: LREAL;(*前次时间|*)
	xReqTestEndVelocity: BOOL;
	lrCurCycleVelVeries: LREAL;(*当前周期速度变化量|*)
	alrInflectionPts_t: ARRAY [1..2] OF LREAL:= [2(0)];(*时间轴上的拐点位置|*)

	xFlag_MotionParamInitialized: BOOL := FALSE;(*运动参数初始化标志|*)

	rMax_a_Coeff: REAL:=1.5;
	rS_AccDecTime_Coeff:REAL;(*S加减速时间-加速占的比例*)
	rAux_enc_vel_Temp:REAL;
	rTemp_Compera_Vel: REAL := 0.000016;
	fbTRIG_ArrivedTOtar: R_TRIG;
	lrFinalVelocity : LREAL;
	rAux_enc_vel : REAL;
END_VAR
{IMPLEMENTATION}
o_xEno:= i_xEn;
o_iErNo:= 0;
(*
IF i_bySTime_AtLeast=0 THEN
	i_bySTime_AtLeast:=10;
END_IF
*)
IF i_rGirth_Master=0 THEN
	i_rGirth_Master:= 0.5;
END_IF
IF i_xEn THEN
	IF
		i_iMsCycle_Motion>0 AND
		i_lrTimeSec_SBegin>0 AND
		i_lrTimeSec_SEnd>0 THEN
		//在这里处理速度到位清标志动作2023.8.17.210154

		IF NOT (i_piTimeSec_AccDec_AllTheWay^(*i_pstStGrpParam^.iTimeSec_AccDec_AllTheWay*)>0
			AND (*i_pstStGrpParam^.lrVel_Max*)i_rVel_Max>0) THEN
			o_iErNo:= -2;
			RETURN;
		END_IF
		fbTRIG_ArrivedTOtar(CLK:=i_pxFlag_ArrivedToTargetVel^);
		IF fbTRIG_ArrivedTOtar.Q THEN
			o_diVel_Virtual_Tar:= REAL_TO_DINT(ABS(i_rAux_enc_vel));
			o_lrMax_a_S_pos:= 1;
			o_lrTime_S:= 0;
		END_IF
		IF (*i_pstStGrpParam^.xFlag_ArrivedToTargetVel*)i_pxFlag_ArrivedToTargetVel^ OR i_xReCalc_Target THEN(*速度到位|*)
			xFlag_MotionParamInitialized:= FALSE;
			o_iErNo:= -3;
			RETURN;
		END_IF

		IF NOT xFlag_MotionParamInitialized THEN(*未初始化就在这里初始化1次|*)
			xFlag_MotionParamInitialized:= TRUE;
			(*平均加速度(m/min/s)|*)
			lrAve_a:= (*i_pstStGrpParam^.l*)i_rVel_Max/INT_TO_LREAL(i_piTimeSec_AccDec_AllTheWay^);
			(*速度变化量|*)
			lrVel_delta:= (*i_pstStGrpParam^.lrFinalVelocity*)i_rFinalVelocity-i_prVel_Cur^(*i_pstStGrpParam^.lrVel_Cur*);

			(*按照平均加速度算出该段速度变化所需要的时间\
			/*由于时间是绝对量\不能出现负值|*)
(*			i_pstStGrpParam^.lrAccDecTime_ThisTime*)
			i_prAccDecTime_ThisTime^:= LREAL_TO_REAL(ABS(lrVel_delta/lrAve_a));

			IF lrVel_delta<0 THEN
				lrAve_a:= -lrAve_a;

			(*2018.11.26.184729|niu.j|判断如果10米印刷停机到10米空转时，
				当前速度等于目标速度导致有加速度计算，直接输出速度到位标志
				速度变化量为0时直接退出，防止rAccDecTime_ThisTime=0,导致除0*)
			ELSIF lrVel_delta=0 THEN
				i_pxFlag_ArrivedToTargetVel^:= TRUE;
				RETURN;
			ELSE;
			END_IF
			(*2022.4.21.163408 增加了自动加减速曲线选择|*)
			(*自动加减速曲线选择|默认 按照最大直线加速度进行s处理-
									 1：按照直线加速时间进行s处理-不限制最大加速度
									 2：按照直线加速时间进行s处理-限制最大加速度
									 3：按照直线加速时间全程s处理-
									 4: 和默认处理方式接近|增加了至少10s的s加减速处理|2022.8.9.091924*)
			rS_AccDecTime_Coeff:= LREAL_TO_REAL(i_lrTimeSec_SBegin/(i_lrTimeSec_SBegin+i_lrTimeSec_SEnd));
			IF i_byAutoAccDecCurve=1 THEN(*按照直线加速时间进行s处理-不限制最大加速度*)
				i_prAccDecTime_ThisTime^:= i_prAccDecTime_ThisTime^;

				IF i_prAccDecTime_ThisTime^>(i_lrTimeSec_SBegin+i_lrTimeSec_SEnd) THEN(*梯形|*)
					iNum_InflectionPts:= 2;
					(*平均加速度(m/min/s)|*)
					IF i_prAccDecTime_ThisTime^*2<>i_lrTimeSec_SBegin+i_lrTimeSec_SEnd THEN
						lrMax_a_S:= 2*lrVel_delta/(2*i_prAccDecTime_ThisTime^-i_lrTimeSec_SBegin-i_lrTimeSec_SEnd);
					END_IF

					lrJerk_SBegin:= lrMax_a_S/i_lrTimeSec_SBegin;
					lrJerk_SEnd:= lrMax_a_S/i_lrTimeSec_SEnd;
					alrInflectionPts_t[1]:= i_lrTimeSec_SBegin;
					alrInflectionPts_t[2]:= i_prAccDecTime_ThisTime^-i_lrTimeSec_SEnd;
				ELSE(*三角形*)
					iNum_InflectionPts:= 1;
					(*平均加速度(m/min/s)|*)
					IF i_prAccDecTime_ThisTime^<>0 THEN
						lrMax_a_S:= 2*lrVel_delta/(i_prAccDecTime_ThisTime^);
					END_IF

					alrInflectionPts_t[1]:= ABS(i_prAccDecTime_ThisTime^*(rS_AccDecTime_Coeff));
					alrInflectionPts_t[2]:= ABS(i_prAccDecTime_ThisTime^*(1-rS_AccDecTime_Coeff));
					lrJerk_SBegin:= lrMax_a_S/alrInflectionPts_t[1];
					lrJerk_SEnd:= lrMax_a_S/alrInflectionPts_t[2];
				END_IF

			ELSIF i_byAutoAccDecCurve=2 THEN(*按照直线加速时间进行s处理-限制最大加速度|这中情况下s加减速时间会变*)
				i_prAccDecTime_ThisTime^:= i_prAccDecTime_ThisTime^;
				(*在不修改s加减速时间计算最大平均加速度(m/min/s)|*)
				IF i_prAccDecTime_ThisTime^>(i_lrTimeSec_SBegin+i_lrTimeSec_SEnd) THEN(*梯形|*)
					IF i_prAccDecTime_ThisTime^*2>i_lrTimeSec_SBegin+i_lrTimeSec_SEnd THEN
						lrMax_a_S:= 2*lrVel_delta/(2*i_prAccDecTime_ThisTime^-i_lrTimeSec_SBegin-i_lrTimeSec_SEnd);
					END_IF
				ELSE
					(*重新计算平均加速度(m/min/s)|*)
					IF i_prAccDecTime_ThisTime^<>0 THEN
						lrMax_a_S:= 2*lrVel_delta/(i_prAccDecTime_ThisTime^);
					END_IF
				END_IF

				IF ABS(lrAve_a)*rMax_a_Coeff<ABS(lrMax_a_S) THEN(*超过了我限制的最大加速度-按照最大加速度处理
													我就需要重新计算s加减速时间*)
					lrMax_a_S:=lrAve_a*rMax_a_Coeff;(*最大加速度为直线加速度的倍数*)

					(*重新计算s时间*)
					i_lrTimeSec_SBegin:=2*(i_prAccDecTime_ThisTime^-ABS(lrVel_delta/lrMax_a_S))*rS_AccDecTime_Coeff;
					i_lrTimeSec_SEnd:=2*(i_prAccDecTime_ThisTime^-ABS(lrVel_delta/lrMax_a_S))*(1-rS_AccDecTime_Coeff);
				END_IF

				IF i_prAccDecTime_ThisTime^>(i_lrTimeSec_SBegin+i_lrTimeSec_SEnd) THEN(*梯形|*)
					iNum_InflectionPts:= 2;

					lrJerk_SBegin:= lrMax_a_S/i_lrTimeSec_SBegin;
					lrJerk_SEnd:= lrMax_a_S/i_lrTimeSec_SEnd;
					alrInflectionPts_t[1]:= i_lrTimeSec_SBegin;
					alrInflectionPts_t[2]:= i_prAccDecTime_ThisTime^-i_lrTimeSec_SEnd;
				ELSE(*三角形*)
					iNum_InflectionPts:= 1;

					alrInflectionPts_t[1]:= ABS(i_prAccDecTime_ThisTime^*(rS_AccDecTime_Coeff));
					alrInflectionPts_t[2]:= ABS(i_prAccDecTime_ThisTime^*(1-rS_AccDecTime_Coeff));
					lrJerk_SBegin:= lrMax_a_S/alrInflectionPts_t[1];
					lrJerk_SEnd:= lrMax_a_S/alrInflectionPts_t[2];
				END_IF

			ELSIF i_byAutoAccDecCurve=3 THEN(*按照直线加速时间全程s处理*)
				(*三角形*)
				iNum_InflectionPts:= 1;
				(*平均加速度(m/min/s)|*)
				IF i_prAccDecTime_ThisTime^<>0 THEN
					lrMax_a_S:= 2*lrVel_delta/(i_prAccDecTime_ThisTime^);
				END_IF

				alrInflectionPts_t[1]:= ABS(i_prAccDecTime_ThisTime^*(rS_AccDecTime_Coeff));
				alrInflectionPts_t[2]:= ABS(i_prAccDecTime_ThisTime^*(1-rS_AccDecTime_Coeff));
				lrJerk_SBegin:= lrMax_a_S/alrInflectionPts_t[1];
				lrJerk_SEnd:= lrMax_a_S/alrInflectionPts_t[2];
			ELSIF i_byAutoAccDecCurve=4 THEN(*和默认处理方式接近|增加了至少10s的s加减速处理|2022.8.9.091924*)
				IF i_xFlag_Print THEN(*增加印刷标志|印刷状态和空转匀墨使用不同加速逻辑|2022.11.06.104252*)
					(*屏蔽之前前后加相等时间的S曲线加速方式|改为前后加不同时间的方式|2023.03.02.112443*)
					(*
						iNum_InflectionPts:=2;(*还是使用T形方式|本次时间前后+i_bySTime_AtLeast时间s*)
						lrMax_a_S:= lrAve_a*i_pstStGrpParam^.lrAccDecTime_ThisTime/(i_pstStGrpParam^.lrAccDecTime_ThisTime+i_bySTime_AtLeast);(*计算最大的加速度*)

						i_pstStGrpParam^.lrAccDecTime_ThisTime:= i_pstStGrpParam^.lrAccDecTime_ThisTime+i_bySTime_AtLeast*2;
						lrJerk_SBegin:= lrMax_a_S/i_bySTime_AtLeast;
						lrJerk_SEnd:= lrMax_a_S/i_bySTime_AtLeast;
						alrInflectionPts_t[1]:= i_bySTime_AtLeast;
						alrInflectionPts_t[2]:= i_pstStGrpParam^.lrAccDecTime_ThisTime-i_bySTime_AtLeast;
	(*2022.12.7.170336@liu
					END_IF
	*)
					*)
						iNum_InflectionPts:=2;(*还是使用T形方式|*)
						(*使用前后不同的S加速时间|2023.03.02.113109|*)
						lrMax_a_S:=2*lrVel_delta/(i_lrTimeSec_SBegin+i_lrTimeSec_SEnd+
									2*i_prAccDecTime_ThisTime^);

						i_prAccDecTime_ThisTime^:= LREAL_TO_REAL(i_prAccDecTime_ThisTime^+i_lrTimeSec_SBegin+i_lrTimeSec_SEnd);
						lrJerk_SBegin:= lrMax_a_S/i_lrTimeSec_SBegin;
						lrJerk_SEnd:= lrMax_a_S/i_lrTimeSec_SEnd;
						alrInflectionPts_t[1]:= i_lrTimeSec_SBegin;
						alrInflectionPts_t[2]:= i_prAccDecTime_ThisTime^-i_lrTimeSec_SEnd;
				ELSE(*使用默认加速方式|2022.11.06.104353*)
					(*平均加速度(m/min/s)|*)
					IF i_prAccDecTime_ThisTime^*2>(i_lrTimeSec_SBegin+i_lrTimeSec_SEnd) THEN(*梯形|*)
						iNum_InflectionPts:= 2;
						i_prAccDecTime_ThisTime^:= LREAL_TO_REAL(i_prAccDecTime_ThisTime^+i_lrTimeSec_SBegin/2.0+i_lrTimeSec_SEnd/2.0);
						lrMax_a_S:= lrAve_a;
						lrJerk_SBegin:= lrMax_a_S/i_lrTimeSec_SBegin;
						lrJerk_SEnd:= lrMax_a_S/i_lrTimeSec_SEnd;
						alrInflectionPts_t[1]:= i_lrTimeSec_SBegin;
						alrInflectionPts_t[2]:= i_prAccDecTime_ThisTime^-i_lrTimeSec_SEnd;
					ELSE(*三角形*)
						iNum_InflectionPts:= 1;
						i_prAccDecTime_ThisTime^:= i_prAccDecTime_ThisTime^*2;
						lrMax_a_S:= lrAve_a;
						alrInflectionPts_t[1]:= i_prAccDecTime_ThisTime^/2;
						alrInflectionPts_t[2]:= i_prAccDecTime_ThisTime^/2;
						lrJerk_SBegin:= lrMax_a_S/alrInflectionPts_t[1];
						lrJerk_SEnd:= lrMax_a_S/alrInflectionPts_t[2];
					END_IF
				END_IF

			ELSE(*默认*)
				(*平均加速度(m/min/s)|*)
				IF i_prAccDecTime_ThisTime^*2>(i_lrTimeSec_SBegin+i_lrTimeSec_SEnd) THEN(*梯形|*)
					iNum_InflectionPts:= 2;
					i_prAccDecTime_ThisTime^:= LREAL_TO_REAL(i_prAccDecTime_ThisTime^+i_lrTimeSec_SBegin/2.0+i_lrTimeSec_SEnd/2.0);
					lrMax_a_S:= lrAve_a;
					lrJerk_SBegin:= lrMax_a_S/i_lrTimeSec_SBegin;
					lrJerk_SEnd:= lrMax_a_S/i_lrTimeSec_SEnd;
					alrInflectionPts_t[1]:= i_lrTimeSec_SBegin;
					alrInflectionPts_t[2]:= i_prAccDecTime_ThisTime^-i_lrTimeSec_SEnd;
				ELSE(*三角形*)
					iNum_InflectionPts:= 1;
					i_prAccDecTime_ThisTime^:= i_prAccDecTime_ThisTime^*2;
					lrMax_a_S:= lrAve_a;
					alrInflectionPts_t[1]:= i_prAccDecTime_ThisTime^/2;
					alrInflectionPts_t[2]:= i_prAccDecTime_ThisTime^/2;
					lrJerk_SBegin:= lrMax_a_S/alrInflectionPts_t[1];
					lrJerk_SEnd:= lrMax_a_S/alrInflectionPts_t[2];
				END_IF
			END_IF

			lrCurr_t:= 0;
			lrPrev_t:= 0;
			//2023.8.17.210752在这里输出一下目标速度和加速度减速度
			//o_iVel_Virtual_Tar:= REAL_TO_INT(i_rFinalVelocity*GC_LRMOTORPPR/1.5/60.0/1000.0);
			//o_lrMax_a_S_pos:= lrMax_a_S*GC_LRMOTORPPR/60.0/1000.0/1000.0;
(*
////////////////////////////////////////////////////////////////////////////////////////////////////////////////////////////////////
			IF i_xFlag_ManuDec OR i_xFlag_EStoping(*2023.08.28.193725*)
				OR i_xFlag_Stoping OR
				i_xFlag_FastStoping THEN(* OR(*手动减速和急停/停机/快速停止中采用直线减速|*)
				(*2023.3.2.164553 空转自动减速也使用直线减速*)
				(i_xFlag_AutoDec AND i_xflag_ink) THEN*)
					o_iVel_Virtual_Tar:= REAL_TO_INT(i_rFinalVelocity*GC_LRMOTORPPR/1.5/60.0/1000.0);
					o_lrMax_a_S_pos:= lrAve_a*GC_LRMOTORPPR/1.5/60.0/1000.0/1000.0;
					o_lrTime_S := 0;
			ELSIF i_xFlag_ManuAcc OR
				i_xFlag_InkAccing (*OR(*手动加速/空转加速用手动直线加速|*)
				(*2023.3.2.164553 空转自动加速使用直线加速*)
				(i_xFlag_AutoAcc AND i_xflag_ink)*) THEN
					o_iVel_Virtual_Tar:= REAL_TO_INT(i_rFinalVelocity*GC_LRMOTORPPR/1.5/60.0/1000.0);
					o_lrMax_a_S_pos:= lrAve_a*GC_LRMOTORPPR/1.5/60.0/1000.0/1000.0;
					o_lrTime_S := 0;
			ELSIF i_xFlag_AutoAcc  OR(*自动加速或空转加速|*)
				i_xFlag_AutoDec OR (*2023.3.2.164553 空转自动减速也使用直线减速*)
				(i_xFlag_AutoDec AND i_xflag_ink) THEN(*自动减速或默认停机|*)
					o_iVel_Virtual_Tar:= REAL_TO_INT(i_rFinalVelocity*GC_LRMOTORPPR/1.5/60.0/1000.0);
					o_lrMax_a_S_pos:= lrMax_a_S*GC_LRMOTORPPR/1.5/60.0/1000.0/1000.0;
					o_lrTime_S := alrInflectionPts_t[1];
			END_IF
*)
////////////////////////////////////////////////////////////////////////////////////////////////////////////////////////////////////
		//2023.10.19.142926
			IF i_xFlag_ManuDec OR i_xFlag_EStoping(*2023.08.28.193725*)
				OR i_xFlag_Stoping OR
				i_xFlag_FastStoping OR(*手动减速和急停/停机/快速停止中采用直线减速|*)
				(*2023.3.2.164553 空转自动减速也使用直线减速*)
				(i_xFlag_AutoDec AND (i_xflag_ink OR i_byAutoAccDecCurve=5)) THEN
					o_diVel_Virtual_Tar:= LREAL_TO_DINT(i_rFinalVelocity*GC_LRMOTORPPR/i_rGirth_Master/60.0/1000.0);
					o_lrMax_a_S_pos:= lrAve_a*GC_LRMOTORPPR/i_rGirth_Master/60.0/1000.0/1000.0;
					o_lrTime_S := 0;
			ELSIF i_xFlag_ManuAcc OR
				i_xFlag_InkAccing OR(*手动加速/空转加速用手动直线加速|*)
				(*2023.3.2.164553 空转自动加速使用直线加速*)
				(i_xFlag_AutoAcc AND (i_xflag_ink OR i_byAutoAccDecCurve=5)) THEN
					o_diVel_Virtual_Tar:= LREAL_TO_DINT(i_rFinalVelocity*GC_LRMOTORPPR/i_rGirth_Master/60.0/1000.0);
					o_lrMax_a_S_pos:= lrAve_a*GC_LRMOTORPPR/i_rGirth_Master/60.0/1000.0/1000.0;
					o_lrTime_S := 0;
			ELSIF i_xFlag_AutoAcc  OR(*自动加速或空转加速|*)
				i_xFlag_AutoDec THEN(*自动减速或默认停机|*)
					o_diVel_Virtual_Tar:= LREAL_TO_DINT(i_rFinalVelocity*GC_LRMOTORPPR/i_rGirth_Master/60.0/1000.0);
					o_lrMax_a_S_pos:= lrMax_a_S*GC_LRMOTORPPR/i_rGirth_Master/60.0/1000.0/1000.0;
					o_lrTime_S := alrInflectionPts_t[1];
			END_IF
		END_IF
//bai.zy | 2024.01.16.103002 | 重新判断标志

		rAux_enc_vel_Temp:= LREAL_TO_REAL(ABS(i_rAux_enc_vel)*1000.0*60.0*i_rGirth_Master/GC_LRMOTORPPR);
		i_prVel_Cur^:= rAux_enc_vel_Temp;
		rAux_enc_vel:= ABS(i_rAux_enc_vel);
		lrFinalVelocity := LREAL_TO_DINT(i_rFinalVelocity*GC_LRMOTORPPR/i_rGirth_Master/60.0/1000.0);

		IF i_iIdGSE=GSE_ACCING OR
			i_iIdGSE=GSE_DECING THEN

			IF i_xFlag_ManuDec OR i_xFlag_EStoping
				OR i_xFlag_Stoping OR
				i_xFlag_FastStoping OR(*手动减速和急停/停机/快速停止中采用直线减速|*)
				(*2023.3.2.164553 空转自动减速也使用直线减速*)
				(i_xFlag_AutoDec AND (i_xflag_ink OR i_byAutoAccDecCurve=5)) THEN
				lrCurCycleVelVeries:= lrAve_a*(INT_TO_LREAL(i_iMsCycle_Motion)/1000);
				IF rAux_enc_vel > lrFinalVelocity + rTemp_Compera_Vel(*i_prVel_Cur^>i_rFinalVelocity+rTemp_Compera_Vel*) THEN
					i_pxFlag_Decing^:= TRUE;
					i_pxFlag_Accing^:= FALSE;
				ELSE
					i_pxFlag_Decing^:= FALSE;
					i_pxFlag_Accing^:= FALSE;
					i_prVel_Cur^:= i_rFinalVelocity;
//2023.8.17.213343到目标速度后，把目标速度再设置一次-为了防止手自动加速过程中停下并且速度同步
					o_diVel_Virtual_Tar:= LREAL_TO_DINT(i_rFinalVelocity*GC_LRMOTORPPR/i_rGirth_Master/60.0/1000.0);
					i_pxFlag_ArrivedToTargetVel^:= TRUE;
				END_IF
			(*2018.10.5.133955 | niu.j | 空转加速采用直线加速*)
			ELSIF i_xFlag_ManuAcc OR
				i_xFlag_InkAccing OR(*手动加速/空转加速用手动直线加速|*)
				(*2023.3.2.164553 空转自动加速使用直线加速*)
				(i_xFlag_AutoAcc AND (i_xflag_ink OR i_byAutoAccDecCurve=5)) THEN

				IF rAux_enc_vel < lrFinalVelocity-rTemp_Compera_Vel(*i_prVel_Cur^<i_rFinalVelocity-rTemp_Compera_Vel *)THEN
					i_pxFlag_Decing^:= FALSE;
					i_pxFlag_Accing^:= TRUE;
				ELSE
					i_pxFlag_Decing^:= FALSE;
					i_pxFlag_Accing^:= FALSE;
					i_prVel_Cur^:= i_rFinalVelocity;
					o_diVel_Virtual_Tar:= LREAL_TO_DINT(i_rFinalVelocity*GC_LRMOTORPPR/i_rGirth_Master/60.0/1000.0);
					i_pxFlag_ArrivedToTargetVel^:= TRUE;
				END_IF
			ELSIF i_xFlag_AutoAcc  OR(*自动加速或空转加速|*)
				i_xFlag_AutoDec THEN(*自动减速或默认停机|*)
				IF (((i_xFlag_AutoAcc OR i_xFlag_InkAccing) AND
						rAux_enc_vel < lrFinalVelocity-rTemp_Compera_Vel) (*i_prVel_Cur^<i_rFinalVelocity-rTemp_Compera_Vel) *)OR
					((i_xFlag_AutoDec OR i_xFlag_Stoping OR i_xFlag_FastStoping) AND
						rAux_enc_vel > lrFinalVelocity+rTemp_Compera_Vel))(*i_prVel_Cur^>i_rFinalVelocity+rTemp_Compera_Vel)) *)THEN

					IF i_xFlag_AutoAcc OR i_xFlag_InkAccing THEN
						i_pxFlag_Accing^:= TRUE;
						i_pxFlag_Decing^:= FALSE;
					ELSE
						i_pxFlag_Accing^:= FALSE;
						i_pxFlag_Decing^:= TRUE;
					END_IF
				ELSE
					i_pxFlag_Decing^:= FALSE;
					i_pxFlag_Accing^:= FALSE;
					i_pxFlag_ArrivedToTargetVel^:= TRUE;
					(*2018.8.15.095720 :| niu.j | 到目标速度后，当前速度赋值为目标速度*)
					i_prVel_Cur^:= i_rFinalVelocity;
					o_diVel_Virtual_Tar:= LREAL_TO_DINT(i_rFinalVelocity*GC_LRMOTORPPR/i_rGirth_Master/60.0/1000.0);
				END_IF
			END_IF

		END_IF

	ELSE
		o_iErNo:= -1;(*Bad parameters|*)
	END_IF
END_IF
